      slope = computeSlope(rawRange, scaledRange)
      intercept = computeIntercept(slope, rawRange, scaledRange)
      scaledValue = slope * value + intercept
      return clipScaledValue(scaledValue, scaledRange)
  end

  def limit(value, range):
      return scale(value, range, range)
  end


  rq_init_comm_if_connected(9, "1")
  rq_init_comm_if_connected(2, "2")
  rq_init_comm_if_connected(3, "3")
  rq_init_comm_if_connected(4, "4")
  rq_print_connected_grippers()
  rq_gripper_communication_thread = run rq_gripper_communication()
  set_closed_norm(97.6470588235294, 1)
  set_open_norm(1.1764705882352942, 1)
  set_closed_mm(0.0, 1)
  set_open_mm(53.0, 1)
  set_closed_norm(100.0, 2)
  set_open_norm(0.0, 2)
  set_closed_mm(0.0, 2)
  set_open_mm(50.0, 2)
  set_closed_norm(100.0, 3)
  set_open_norm(0.0, 3)
  set_closed_mm(0.0, 3)
  set_open_mm(50.0, 3)
  set_closed_norm(100.0, 4)
  set_open_norm(0.0, 4)
  set_closed_mm(0.0, 4)
  set_open_mm(50.0, 4)
  rq_current_limit_enabled = False
  while(not rq_gripper_communication_thread_started):
      sync()
  end
  # end: URCap Installation Node
  # begin: URCap Installation Node
  #   Source: OPC UA, 2.0.2, Rocketfarm AS
  #   Type: OPC UA
  global opcua_daemon = rpc_factory("xmlrpc", "http://127.0.0.1:40409/RPC2")
  def opcua_client_connect(address):
  return opcua_daemon.client_connect(address)
  end
  def opcua_client_get_id(client_name):
  return opcua_daemon.client_get_id(client_name)
  end
  def opcua_client_try_connect(client_id):
  opcua_result = False
  if (opcua_daemon.client_connect(client_id)):
  sleep(0.01)
  opcua_result = opcua_daemon.client_is_connected(client_id)
  opcua_retry = 10
  while ( (not opcua_result) and (opcua_retry > 0) ):
  sleep(0.1)
  opcua_result = opcua_daemon.client_is_connected(client_id)
  opcua_retry = opcua_retry - 1
  end
  end
  return opcua_result
  end
  def opcua_client_disconnect(client_id):
  return opcua_daemon.client_disconnect(client_id)
  end
  def opcua_client_is_connected(client_id):
  return opcua_daemon.client_is_connected(client_id)
  end
  def opcua_client_read_byid(client_id, namespace_id, variable_id):
  return opcua_daemon.client_read_variable_by_id(client_id, namespace_id, variable_id)
  end
  def opcua_client_read_byname(client_id, namespace_id, variable_name):
  return opcua_daemon.client_read_variable_by_name(client_id, namespace_id, variable_name)
  end
  def opcua_client_write_byid(client_id, namespace_id, variable_id, variable_value):
  return opcua_daemon.client_write_variable_by_id(client_id, namespace_id, variable_id, variable_value)
  end
  def opcua_client_write_byname(client_id, namespace_id, variable_name, variable_value):
  return opcua_daemon.client_write_variable_by_name(client_id, namespace_id, variable_name, variable_value)
  end
  def opcua_client_last_error(client_id):
  return opcua_daemon.client_get_last_error(client_id)
  end
  def opcua_server_read_byname(variable_name):
  return opcua_daemon.server_read_variable_by_name(variable_name)
  end
  def opcua_server_write_byname(variable_name, variable_value):
  return opcua_daemon.server_write_variable_by_name(variable_name, variable_value)
  end
  def opcua_server_last_error():
  return opcua_daemon.server_get_last_error()
  end
  def opcua_error_to_string(errorCode):
  return opcua_daemon.error_code_to_string(errorCode)
  end
  # end: URCap Installation Node
  global AMR_Position=struct(position_identifier=0, x1=0, x2=0, y1=0, y2=0, theta1=0, theta2=0)
  global CAM_Pose=p[0,0,0,0,0,0]
  global CAM_Relation=""
  global CMD_Abort=  False
  global CMD_Clear=  False
  global CMD_Reset=  False
  global CMD_Start=  False
  global CMD_Suspend=  False
  global CMD_Unhold=  False
  global CMD_Unsuspend=  False
  global CNT_Rack_Output=0
  global FNC_Freedrive=  False
  global PRC_TubCounter=0
  global STP=0
  global easyPickCount=0
  global easyPickCount_4=0
  global easyPickCount_6=0
  global easyPickNoObj=0
  global easyPickNoObj_4=0
  global easyPickNoObj_6=0
  global easyPickParts=0
  global easyPickParts_4=0
  global easyPickParts_6=0
  global Container_mid_1_p=p[-.379239199143, -.127191311915, .299999999998, .000000000046, -.000000000021, -1.247199999994]
  global Container_mid_1_q=[-2.477408934449926, -1.2969853503591224, -1.875639182904262, -1.539621866126728, 1.5731943360401213, -2.8009955944022717]
  global Container_capt_p=p[-.525590029047, .407247642794, .411588185841, -.000000000107, .000000000065, -2.896148821900]
  global Container_capt_q=[-3.5968351615224767, -2.0050156108707204, -0.8176271154495112, -1.8895759482008394, 1.5730967555598792, -2.2743681102957645]
  global Waypoint_51_p=p[-.335468094724, -.217855817953, .299999999998, .000000000047, -.000000000014, -.994837065669]
  global Waypoint_51_q=[-2.2250460001249586, -1.2969853503591224, -1.875639182904262, -1.539621866126728, 1.573194336040121, -2.800995594402271]
  global Waypoint_65_p=p[-.380578560601, .136229906820, .300065486591, .002668209125, -.001950299791, -1.918285884015]
  global Waypoint_65_q=[-3.1484482924090784, -1.309784547691681, -1.8656262159347534, -1.5396564540318032, 1.5732260942459106, -2.8009706179248255]
  global Waypoint_86_p=p[-.610891912545, .328076512140, .154928874949, -.144389774448, 2.158207980619, -2.101916875088]
  global Waypoint_86_q=[-3.0298424402820032, -2.1616608105101527, -1.770405888557434, -1.8800016842284144, -0.04927570024599248, -0.4936583677874964]
  global Waypoint_16_p=p[-.530358413935, .418971000515, -.109643658887, -.463059997969, 2.087871459122, -2.058033430549]
  global Waypoint_16_q=[-3.2300904432879847, -2.6409207783141078, -1.877760410308838, -1.6937691173949183, -0.43063193956484014, 0.029483795166015625]
  global Waypoint_87_p=p[-.459488806274, .188986755628, .171097942578, -.348072585494, -2.059579317749, 2.019661285019]
  global Waypoint_87_q=[-2.790591303502218, -2.152559896508688, -1.6884642839431763, -2.469414850274557, 0.6884214878082275, 0.021232735365629196]
  global Waypoint_89_p=p[-.261886355761, -.111669623901, .131097242659, -1.173634433322, -1.227274747052, 1.193766216763]
  global Waypoint_89_q=[-2.672995464666928, -2.175407175402028, -1.7617490112425536, -2.338843663300132, 2.030865036219133, 0.036428578240585985]
  global Waypoint_90_p=p[-.269165142951, -.108082457315, .026677271969, -1.173634433324, -1.227274747052, 1.193766216762]
  global Waypoint_90_q=[-2.6853380119023815, -2.380020912479904, -1.7522585114443245, -2.1436252765786143, 2.018787725064888, 0.03659425986402358]
  global Waypoint_88_p=p[-.617446503519, .392270291627, .170489198955, -.224010410006, -2.066036920971, 2.088909130040]
  global Waypoint_88_q=[-3.1488035953258766, -2.4221038789008897, -1.1666724558911366, -2.618578428321003, 0.2380794033913185, -0.04528854192806264]
  global Waypoint_94_p=p[-.452978066378, .173533334300, .109390198136, -.002578830757, -2.196586508502, 2.177068753404]
  global Waypoint_94_q=[-2.6674557574892073, -2.1212895090252317, -1.967198705482553, -2.208419381150989, 0.5117897724834828, 0.04481344519449531]
  global Waypoint_93_p=p[-.596468537907, .142788156334, .105779109453, -.673355127215, 1.831389627653, -1.853156743314]
  global Waypoint_93_q=[-2.6921545586066635, -2.073966887503291, -2.065600898968258, -2.154852607781155, -0.22224352987151796, 0.042304121657345886]
  global Waypoint_95_p=p[-.605386387448, -.069660570533, .218481828695, .000812734400, .006677866481, -1.958478278110]
  global Waypoint_95_q=[-2.8029143834677903, -1.8400819882842256, -1.544169955118452, -1.327224466208456, 1.5676652012497132, -2.4155226342256775]
  global Waypoint_13_p=p[-.479450777041, .284140798427, .125270103493, -.276792173670, 2.098433187455, -2.121256516887]
  global Waypoint_13_q=[-2.8915050665484827, -1.9549266300597132, -2.2318272590637207, -1.6654960117735804, 0.020810842514038086, -0.4019392172442835]
  global Waypoint_70_p=p[-.472820924464, .292439826304, .207418370234, -.259787347864, -2.053484648504, 2.070709755662]
  global Waypoint_70_q=[-2.969927421603815, -2.07168115810532, -1.6835546062719366, -2.4953958198513964, 0.4489790927922641, -0.005578998612037367]
  global Waypoint_2_p=p[-.312961047461, -.152991312519, .223609826854, -.745314530454, -1.713873240489, 1.673341715282]
  global Waypoint_2_q=[-2.3560472170459192, -2.183784624139303, -1.4583134651184082, -2.6435262165465296, 1.6522362232208252, 0.043451953679323196]
  global Waypoint_3_p=p[-.113749865836, -.390110151572, .317307487562, -.519383711706, -.839884211339, 1.756868173041]
  global Waypoint_3_q=[-1.8909733931170862, -1.720626016656393, -1.5115610361099243, -2.1240560017027796, 2.1809096336364746, 0.7227501273155212]
  global Waypoint_15_p=p[.029144035010, -.436802470887, .327885032028, -.521560953301, -.623641814548, 1.862659450154]
  global Waypoint_15_q=[-1.564817253743307, -1.556895188321807, -1.6826975345611572, -1.6944714985289515, 2.2362685203552246, 1.117417335510254]
  global Waypoint_14_p=p[.068712235638, -.569419545175, .285215357659, -.679242949116, -.712065334485, 1.394044574094]
  global Waypoint_14_q=[-1.5731792953485346, -1.8029235103747094, -1.6781008808776736, -1.2218450646111982, 2.4719572998240125, 1.6394218026856375]
  global Waypoint_4_p=p[-.047220457210, -.557624911767, .136370962514, -.679242949107, -.712065334475, 1.394044574096]
  global Waypoint_4_q=[-1.7740079055958748, -2.0023561428872334, -1.7577251142892676, -1.18903287716154, 2.4487287370345143, 1.322902469273079]
  global Waypoint_25_p=p[.065436479647, -.569388431626, .287820755049, -.679242949185, -.712065334557, 1.394044574070]
  global Waypoint_25_q=[-1.5789263550890595, -1.8020194754825436, -1.6702557537748035, -1.237882536889547, 2.471995808083492, 1.6301087487321393]
  global Waypoint_39_p=p[.137772150180, -.577759956854, .299999999946, .000000000217, -.000000000207, -1.594351842625]
  global Waypoint_39_q=[-1.108978697428574, -1.776486680444405, -1.413737665315093, -1.5218908901738937, 1.5733062372356947, -1.0863866394180182]
  global Waypoint_41_p=p[.074222967010, -.565641640647, .234620140366, -.516884386806, .529223682286, -1.529619060506]
  global Waypoint_41_q=[-0.9596722604286052, -1.8767069964135548, -1.4892746174057256, -1.7813862040292285, 1.0520698599867686, -0.8199687448260349]
  global Waypoint_40_p=p[.039987741677, -.564832865048, .191055405868, -.767560686167, .343136533060, -2.241315728308]
  global Waypoint_40_q=[-1.0070649180116558, -1.8745927522477324, -1.6139175023195245, -1.6337474788493545, 1.032708081143138, -0.11587278312988403]
  global Waypoint_42_p=p[.041363380882, -.564865360786, .192805844739, .278500165520, .624117100927, .762272396553]
  global Waypoint_42_q=[-1.0050718976263102, -1.8744386685524779, -1.609151451954446, -1.6399653140247947, 1.0334006002355505, -3.254032861659603]
  global Waypoint_43_p=p[.041363380886, -.564865360780, .192805844755, .854271020883, .226833028600, 2.453002871494]
  global Waypoint_43_q=[-1.0050567614299233, -1.874341297657562, -1.6092945416026048, -1.6397580431809713, 1.0333661149462194, -5.0371728933995605]
  global Waypoint_44_p=p[.040882892233, -.564854254876, .192193763716, .110913882012, .659173708659, .275719738520]
  global Waypoint_44_q=[-1.0057704811530535, -1.8745207681598055, -1.6107765025572558, -1.637858394640876, 1.033164860873599, -2.7487836132940755]
  global Waypoint_45_p=p[.042647731639, -.564895808997, .194439423694, -.451694728506, .563172064821, -1.343350300184]
  global Waypoint_45_q=[-1.0032860829914387, -1.8741561795270565, -1.6048483308761785, -1.6453689714776623, 1.0342050634514657, -1.06078829880322]
  global Waypoint_46_p=p[.099944144487, -.566244126804, .267342790130, -.451694834765, .563172023386, -1.343350532536]
  global Waypoint_46_q=[-0.9257438092434924, -1.889970530402497, -1.3828165217629076, -1.8916791100652528, 1.0664350961373816, -0.9805910833329659]
  global Waypoint_47_p=p[.099944144444, -.566244126727, .267342790273, -.101742139519, .058679218003, -1.457888523314]
  global Waypoint_47_q=[-1.1112623176383014, -1.729989471869196, -1.5530029871033957, -1.4442770617454777, 1.4670579052775654, -1.2224020460061675]
  global Waypoint_48_p=p[-.136182767566, -.647487115908, .294247768372, -.101742139549, .058679218020, -1.457888523312]
  global Waypoint_48_q=[-1.532196177857717, -1.9115932455375173, -1.2651848069729779, -1.5055651746702665, 1.4703193777418382, -1.646379689188814]
  global Waypoint_49_p=p[-.159024328559, -.641021381179, .047691706070, -.000000000033, -.000000000027, -1.457897102937]
  global Waypoint_49_q=[-1.6098490079965062, -2.1164987141784586, -1.6156631902166785, -0.9800092198841526, 1.573231151532669, -1.722204302767242]
  global Waypoint_50_p=p[-.159024328558, -.641021381151, .291114489351, -.000000000033, -.000000000027, -1.457897102937]
  global Waypoint_50_q=[-1.609190265995684, -1.9426985888940234, -1.2189094859258596, -1.55056435122874, 1.5734384912955113, -1.7235116759964022]
  global Waypoint_53_p=p[-.050111345339, -.357608435610, .335880801283, .034180375734, .020280946727, -.284888945062]
  global Waypoint_53_q=[-1.3262308189700454, -1.2221767968893875, -1.8246061249803773, -1.7046285947349489, 1.567288986353525, -2.612420684434543]
  global Spatula_above_p=p[.240417564690, -.250827350286, .422801778001, .000126133258, .000019566993, -.045497134322]
  global Spatula_above_q=[-0.4110710190165463, -1.2060566172281924, -1.6172668714852705, -1.8889350758294619, 1.573016581809478, -1.9375501213280995]
  global Spatula_pick_p=p[.245838473482, -.255593930771, .230843335453, .000126133133, .000019564704, -.045497134323]
  global Spatula_pick_q=[-0.4194386807260848, -1.1902770326089298, -2.122244212434893, -1.399738227295769, 1.573431592600495, -1.943921578313585]
  global container_start_p=p[.200650292946, -.570238751958, .366326773614, 1.360500828661, .021700128770, 2.681649891414]
  global container_start_q=[-0.7669977765142582, -2.188996679669204, -0.7412727239230232, -2.581362891432544, 1.0193601740278728, 1.1884911920528847]
  global container_wp_1_p=p[.170613637794, -.572150573676, .294509026043, 1.259497117139, -.008270589399, 2.787717865625]
  global container_wp_1_q=[-0.8129253370121727, -2.0726598902108755, -1.0846040680899218, -2.2403146195823957, 1.0281191187839607, 1.0435744211830564]
  global Waypoint_55_p=p[.077280900603, -.567308602990, .212067617714, 1.259497117148, -.008270589399, 2.787717865619]
  global Waypoint_55_q=[-0.9181858327853867, -1.9744793804952083, -1.4540279077890048, -1.9155621911627945, 0.9643238328181578, 0.9457250675800015]
  global Waypoint_56_p=p[.135568164031, -.570867938153, .245215470413, 1.476861317558, -.018269607491, 2.679642659499]
  global Waypoint_56_q=[-0.8259784040282607, -2.108036981522602, -1.2111990877342924, -2.2405969375728745, 0.9451797152137279, 1.125710531287379]
  global Waypoint_74_p=p[.164827890887, -.574638012411, .193751361296, 2.053636896063, -.046507887560, 2.274278266449]
  global Waypoint_74_q=[-0.7657213433975762, -2.450387120010788, -0.9886183070290357, -2.7078095590939375, 0.8831550681477878, 1.5106229631053527]
  global ftr_scoop2_p=p[.194287054614, -.495779761333, .282072128495, -.179029871953, 1.612108092436, -.016025695011]
  global ftr_scoop2_q=[-0.5957383150173561, -2.264100500923713, -1.1936887184643812, -2.8893702964346097, 0.8750688478879766, -1.4109843517598684]
  global aftr_scoo3_p=p[-.289759911340, -.315385007342, .303743796282, .159961590809, 1.627415489603, -.344855744095]
  global aftr_scoo3_q=[-1.3374747909924949, -1.6809733407851706, -1.9857606509106667, -2.713564895186775, 0.5589807453366573, -1.3631067603374376]
  global Waypoint_60_p=p[-.013316432876, -.544772031582, .383371643081, 2.208233379808, .037543335712, 2.097559881761]
  global Waypoint_60_q=[-0.9328326161883087, -2.0999933666355775, -1.1958015693111372, -3.060905141293654, 0.690378518537611, 1.7121940951337198]
  global Waypoint_61_p=p[-.412188693372, -.356446875193, .383371643081, 1.751740964455, -.739956256289, 1.600691174920]
  global Waypoint_61_q=[-1.766185342973321, -2.0999933666355775, -1.1958015693111372, -3.060905141293654, 0.690378518537611, 1.7121940951337198]
  global Waypoint_75_p=p[-.343126484123, -.342779621892, .335357223804, .359429517288, 1.600352990741, -.365083732359]
  global Waypoint_75_q=[-1.517806275013295, -1.8136828056045395, -1.737638081810795, -2.8432599585466436, 0.5149430839716123, -1.4579122147201877]
  global aftr_scoop1_p=p[.138503854266, -.514479969882, .214153672011, -.134825326227, 1.559916297527, -.059196589314]
  global aftr_scoop1_q=[-0.6880464314785328, -2.2689986529709643, -1.3310176475983653, -2.673087158390708, 0.8340516295138949, -1.4557846480003231]
  global After_disp_3_p=p[.125934854156, -.585611107804, .299545938076, .959554236104, -.134386766509, 2.880651774211]
  global After_disp_3_q=[-0.9434480594885066, -2.016473586333989, -1.1036579072158617, -2.096459283015281, 1.1479556364931514, 0.8433331387406042]
  global Waypoint_62_p=p[-.542658707241, -.114281911009, .251261544113, 1.813043609523, -.679411528034, 1.655271622964]
  global Waypoint_62_q=[-2.158300033470912, -1.9418836862428677, -1.8142999147147894, -2.778920736683023, 0.21900622104017292, 1.8983390235012934]
  global Waypoint_63_p=p[.101294795191, -.465376052375, .381756220355, .972633305146, -.158447626639, 2.887199602585]
  global Waypoint_63_q=[-0.8528172446194038, -1.7393709485118478, -1.2544079521837954, -2.2703112963960628, 1.1965892397133469, 0.91867216443391]
  global Start_p=p[-.033064633790, -.365398531763, .389873206922, .000000000001, .000000000001, 2.725785203584]
  global Start_q=[-1.287596562866887, -1.232866726886848, -1.6880113260231102, -1.7912103151657988, 1.5729028131945846, 0.6981423183093938]
  global Waypoint_76_p=p[-.479450777041, .284140798427, .125270103493, -.276792173670, 2.098433187454, -2.121256516887]
  global Waypoint_76_q=[-2.891505066548503, -1.9549266300590151, -2.231827259067863, -1.6654960117542226, 0.020810842514162875, -0.4019392172601952]
  global PowderA_wayp1_p=p[-.472820924474, .292439826233, .207418370237, -.137787250486, 2.177332259632, -2.152029714756]
  global PowderA_wayp1_q=[-2.911134078210732, -1.90240864358569, -1.968768330510411, -2.500365101593811, 0.11427687110891149, 0.0958980389250167]
  global Waypoint_80_p=p[-.303921889165, -.326082520111, .297721580072, -.584846481381, 1.914382606328, -1.960922301253]
  global Waypoint_80_q=[-1.6364180099980672, -2.041258366871811, -1.472153549517767, -2.7572808013122696, 0.9684003593854582, 0.047163023020230455]
  global Decapp_above_p=p[-.013480295948, -.359153355979, .266194408367, -.879653555922, 1.646336924805, -1.709111068605]
  global Decapp_above_q=[-0.9632157249872035, -2.0163405763031657, -1.5968194594157152, -2.6579215719847085, 1.251243398585566, 0.047906446502667066]
  global Decapp_place_p=p[-.013480295848, -.359153356116, .158558645017, -.879653554904, 1.646336919751, -1.709111066446]
  global Decapp_place_q=[-0.9633419174801583, -2.157735564881908, -1.695182597572722, -2.418253553201909, 1.2517436353048952, 0.04819090596102882]
  global Waypoint_78_p=p[-.051450028091, -.519555688329, .365718563414, -1.287302938145, 1.077637394477, -1.218524965834]
  global Waypoint_78_q=[-0.9214276262416012, -1.8899696965062578, -1.4939326452510562, -2.840015661555725, 0.5585157189668353, 0.033997638875617575]
  global Waypoint_81_p=p[-.030847790230, -.346237542439, .241203613248, .000000000000, .000000000000, .000000000000]
  global Waypoint_81_q=[-1.265848516232941, -1.1652881302267932, -2.11003646605462, -1.4369228603041853, 1.573284436504383, -2.835929896730388]
  global Waypoint_79_p=p[-.030847972829, -.346235312674, .229874122470, .000000000000, .000000000000, .000000000000]
  global Waypoint_79_q=[-1.2659333103898618, -1.1699230683425625, -2.1365870669440055, -1.4057372655396474, 1.5732787836040316, -2.8358953794066757]
  global Waypoint_82_p=p[-.031079593487, -.346547394534, .293012696855, -.000011575267, -.000017731224, -.000713984074]
  global Waypoint_82_q=[-1.2664169521879751, -1.1572597700415788, -1.982185304253158, -1.5727862504184884, 1.5732673022058234, -2.83632822711502]
  global Cap_above_p=p[-.163602500478, -.618357694237, .258271116068, .000026793591, -.000032305852, -.969382601663]
  global Cap_above_q=[-1.6181634639269902, -1.896432778341337, -1.3662765317923142, -1.449515114018281, 1.5734416863575176, -2.220489512402157]
  global Cap_Place_p=p[-.153420247224, -.637174247221, .035295616791, .000000000002, -.000000000002, -1.457849918374]
  global Cap_Place_q=[-1.6014084627078784, -2.123124488207292, -1.6429187572395012, -0.946127085055064, 1.573175527437006, -1.7136981844648291]
  global OP_PowderA2_p=p[.009371277507, -.409434369247, .294169017766, -.823281033205, 1.709410851243, -1.698303593897]
  global OP_PowderA2_q=[-0.9994544761745754, -2.1395254572673217, -1.3437567783153916, -2.8143375616690456, 1.2617899549595724, 0.019614613715634555]
  global OP_PowderA_abov_p=p[-.012145216791, -.363335041455, .315325728178, -.777135478411, 1.752984823781, -1.740925591659]
  global OP_PowderA_abov_q=[-1.01634425044037, -2.024785947780374, -1.4658894155189923, -2.8070189735738786, 1.3091674480404514, 0.020022086766872782]
  global OP_PowderA_pick_p=p[-.012145216707, -.363335041590, .179898787547, -.777135478413, 1.752984823781, -1.740925591659]
  global OP_PowderA_pick_q=[-1.0165129229305911, -2.176980100858497, -1.6127054339661555, -2.5080740815244567, 1.3098787614888208, 0.020270375244195882]
  global Tilt_above_p=p[-.111064400266, -.518714782683, .336190805493, -1.186264705469, 1.271052138367, -1.268665700837]
  global Tilt_above_q=[-1.0593782044036235, -1.983218206819794, -1.4684292238819445, -2.8468741750118465, 0.5899608864573523, 0.021166292918283425]
  global Tilt_place_p=p[-.116477368770, -.516998826303, .220965575609, -1.186264705477, 1.271052138372, -1.268665700834]
  global Tilt_place_q=[-1.0667718212381487, -2.0926346913000655, -1.6256300657432945, -2.5807129872023205, 0.5834128338282412, 0.021733786155414034]
  global Waypoint_52_p=p[-.141928460719, -.515782557948, .252798475575, .000000001021, .000000015714, -1.648489523537]
  global Waypoint_52_q=[-1.5865298660227536, -1.6477298798514424, -1.683499112918053, -1.3809236418182405, 1.5732592408189925, -1.5089407655972176]
  global ViaPoint_1_p=p[-.075380379718, -.518346610957, .240267869004, -.308187611455, .314849234097, -1.629298408213]
  global ViaPoint_1_q=[-1.2665498468402658, -1.632968153584656, -1.7466488267795093, -1.4757122352125567, 1.206407674916738, -1.1583391815257933]
  global Waypoint_57_p=p[-.016929050533, -.520720414258, .208138086750, -.566600031366, .578847302089, -1.576463827532]
  global Waypoint_57_q=[-1.0408435604305932, -1.753222942634757, -1.738239877480245, -1.6732057965873945, 0.9875721214075002, -0.8174462985078907]
  global Waypoint_69_p=p[.038244169892, -.523681622326, .270660553693, -.566600038239, .578847306557, -1.576463843233]
  global Waypoint_69_q=[-0.9584046232102423, -1.7662930703212236, -1.5465420531532832, -1.8980111501412296, 1.0250918773452096, -0.7315432464998608]
  global PowA_ScoopA_p=p[.159611615818, -.500668442765, .327719041452, -.697225816707, .808151787064, -1.272841262549]
  global PowA_ScoopA_q=[-0.7052336156646533, -1.9354458065172322, -1.2435429111590262, -2.383130756765686, 0.9889263119369867, -0.6132400042961272]
  global scoop_p=p[.074657261350, -.519131732172, .256549412299, -.011051468192, .988408833954, .005144340905]
  global scoop_q=[-0.8274053586011583, -1.874926877200366, -1.5200461069833828, -2.106983319332074, 0.9002119871547718, -2.116685021101622]
  global Waypoint_71_p=p[.177770645713, -.528015530173, .277526412330, .001909155730, 1.639086158711, -.035491055298]
  global Waypoint_71_q=[-0.6883155724662711, -2.3735431185097156, -1.0244077123914472, -2.9690624372933723, 0.9072837830600953, -1.4995275296364206]
  global Waypoint_83_p=p[.150765656890, -.528941996739, .207349351161, .001909146913, 1.639086162262, -.035491054401]
  global Waypoint_83_q=[-0.715557591216621, -2.395263074398475, -1.1745539289501714, -2.7990107897487184, 0.8808120190924962, -1.4964991406090151]
  global Waypoint_73_p=p[.145083518034, -.526977858919, .266012644295, -.001096606732, 1.243803685484, -.039558884435]
  global Waypoint_73_q=[-0.7315307126590884, -2.1222688412291646, -1.2371995036129686, -2.500626334721838, 0.9062275384215436, -1.820210419506548]
  global aftr_disp4_p=p[.076649091963, -.516683659078, .327659997949, -.089442013925, .747027934620, -.179429504000]
  global aftr_disp4_q=[-0.8729541889129182, -1.7538731498931135, -1.421722565562387, -2.0624433405073983, 1.0093695837082866, -2.1021195561352615]
  global Waypoint_84_p=p[.123174711194, -.515520147762, .377487231436, -.089442013731, .747027928699, -.179429504004]
  global Waypoint_84_q=[-0.8099995125927881, -1.8159482911699527, -1.2110272502558486, -2.243587231698566, 1.0414314296112155, -2.0397317655088933]
  global Waypoint_54_p=p[.127020102667, -.520474555499, .444734866371, -.000000000049, -.000000000029, -.181836163636]
  global Waypoint_54_q=[-1.077914415145683, -1.67713376904155, -1.1559751108552438, -1.8791222047311322, 1.5728513980826264, -2.469046273458339]
  global Waypoint_58_p=p[.222355978426, -.256721511160, .377517216113, .000126133135, .000019564704, -.045497133314]
  global Waypoint_58_q=[-0.4523685080439055, -1.1582470295698233, -1.764486450044644, -1.7895331365539002, 1.573203470967134, -1.9783680221047675]
  global Waypoint_59_p=p[.246090929453, -.257346948962, .334937874481, .002062251865, .085969144325, -.045466267072]
  global Waypoint_59_q=[-0.3993250128175445, -1.229937207675869, -1.8134849075269486, -1.7494730648138157, 1.5434956294817688, -1.9239935269750585]
  global Waypoint_72_p=p[.241373394141, -.257127682308, .280144245911, .002062251870, .085969144324, -.045466267071]
  global Waypoint_72_q=[-0.40453618428666793, -1.2163524390607545, -1.961899201118312, -1.614505550067273, 1.54321918600584, -1.9286199875396806]
  global Waypoint_68_p=p[-.054140750939, -.519225939047, .230771617164, -.396603942010, .405176681937, -1.615073614845]
  global Waypoint_68_q=[-1.1801200722220573, -1.66078878572511, -1.7519948628362751, -1.5321103532497595, 1.1202658922042295, -1.0435495794713274]
  global Waypoint_67_p=p[-.085538600094, -.517926057057, .244809615848, -.265837410279, .271583584295, -1.634720190296]
  global Waypoint_67_q=[-1.3101477871233094, -1.6246275760972235, -1.7396885526482375, -1.4554188629779246, 1.2515887427265664, -1.211612237682651]
  global Waypoint_66_p=p[-.112404525053, -.516834057197, .249908478866, -.145067433961, .148203121183, -1.645288419275]
  global Waypoint_66_q=[-1.4361046238427022, -1.62151199833529, -1.7216739172895004, -1.4033237867418515, 1.391749278833954, -1.3534436213375054]
  global Waypoint_77_p=p[-.029562189306, -.345402935881, .227061086376, -.000128098079, -.000007607820, -.000007077939]
  global Waypoint_77_q=[-1.2613241377464561, -1.168338291946169, -2.144792803677632, -1.3989918632055023, 1.5732473641903764, -2.831248128197144]
  def Sub_Vision_V18():
    $ 672 "Sub_Vision_V18" "noBreak"
    $ 673 "PreSettings"
    $ 674 "CAM_LM_Detected≔ False "
    global CAM_LM_Detected=  False
    $ 675 "CAM_Captures≔0"
    global CAM_Captures=0
    $ 676 "CAM_Pose≔p[0,0,0,0,0,0]"
    global CAM_Pose=p[0,0,0,0,0,0]
    $ 677 "CAM_LM_Refinmnt≔ False "
    global CAM_LM_Refinmnt=  False
    $ 678 "CAM_LM_Refined≔ False "
    global CAM_LM_Refined=  False
    $ 679 "CAM_LM_Deviatn≔p[0,0,0,0,0,0]"
    global CAM_LM_Deviatn=p[0,0,0,0,0,0]
    $ 680 "CAM_LM_ID≔0"
    global CAM_LM_ID=0
    $ 681 "CAM_Done≔ False "
    global CAM_Done=  False
    $ 682 "CAM_CNT_Obj≔0"
    global CAM_CNT_Obj=0
    $ 683 "CAM_Result = []"
    CAM_Result = []
    $ 684 "OBJ_Detected≔ False "
    global OBJ_Detected=  False
    $ 685 "FRM_Reference≔p[0,0,0,0,0,0]"
    global FRM_Reference=p[0,0,0,0,0,0]
    $ 686 "'=========='"
    # '=========='
    $ 687 "Switch Action"
    switch_1 = Action
    $ 688 "Case 13"
    if (13 == switch_1):
    elif (15 == switch_1):
      $ 806 "Case 15"
    elif (131 == switch_1):
      $ 852 "Case 131"
      $ 853 "Read (SensoPart)"
      $ 854 "Action_Info≔'search for landmark'"
      global Action_Info="search for landmark"
      $ 855 "CAM_LM≔CAM_LMs[4]"
      global CAM_LM=CAM_LMs[4]
      $ 856 "CAM_Relation≔CAM_LM.capture_relation"
      global CAM_Relation=CAM_LM.capture_relation
      $ 857 "go to capture pose"
      $ 860 "If ITM_ID≟1 and JIG≟7"
      if (ITM_ID == 1  and  JIG == 7):
        $ 861 "PSE_T≔uLM_Cap_SSRack"
        global PSE_T=uLM_Cap_SSRack
      else:
        $ 862 "ElseIf ITM_ID≟5 and JIG≟7"
        if (ITM_ID == 5  and  JIG == 7):
          $ 863 "PSE_T≔FRM_Cap_SSRack"
          global PSE_T=FRM_Cap_SSRack
        else:
          $ 864 "ElseIf ITM_ID≟13 and JIG≟7"
          if (ITM_ID == 13  and  JIG == 7):
            $ 865 "PSE_T≔FRM_pick_rack_const"
            global PSE_T=p[-0.5568395192387274,0.34423986364170267,0.44698620470146266,-1.0069110132199915E-6,3.378712467497258E-5,-8.002029546773325E-6]
          else:
            $ 866 "ElseIf ITM_ID≟1 and JIG≟15"
            if (ITM_ID == 1 and JIG == 15):
              $ 867 "MoveJ"
              $ 868 "Container_mid_1" "breakAfter"
              movej(get_inverse_kin(Container_mid_1_p, qnear=Container_mid_1_q), a=1.3962634015954636, v=1.0471975511965976, r=0.05)
              $ 869 "Container_capt" "breakAfter"
              movej(get_inverse_kin(Container_capt_p, qnear=Container_capt_q), a=1.3962634015954636, v=1.0471975511965976)
              $ 870 "PSE_T≔FRM_Container_S_const"
              global PSE_T=p[-0.510412665574981,0.40064363362973565,0.41159789496794374,-1.1370875604168537E-5,-3.643547521609506E-6,-2.896122366208473]
            else:
              $ 871 "ElseIf ITM_ID≟1 and JIG≟16"
              if (ITM_ID == 1  and  JIG == 16):
                $ 872 "MoveJ"
                $ 873 "Waypoint_51" "breakAfter"
                movej(get_inverse_kin(Waypoint_51_p, qnear=Waypoint_51_q), a=1.3962634015954636, v=1.0471975511965976, r=0.05)
                $ 876 "PSE_T≔FRM_Container_S_const"
                global PSE_T=p[-0.510412665574981,0.40064363362973565,0.41159789496794374,-1.1370875604168537E-5,-3.643547521609506E-6,-2.896122366208473]
              else:
                $ 877 "ElseIf ITM_ID≟1 and JIG≟17"
                if (ITM_ID == 1  and  JIG == 17):
                  $ 878 "MoveJ"
                  $ 879 "Waypoint_51" "breakAfter"
                  movej(get_inverse_kin(Waypoint_51_p, qnear=Waypoint_51_q), a=1.3962634015954636, v=1.0471975511965976, r=0.05)
                  $ 882 "PSE_T≔FRM_Container_S_const"
                  global PSE_T=p[-0.510412665574981,0.40064363362973565,0.41159789496794374,-1.1370875604168537E-5,-3.643547521609506E-6,-2.896122366208473]
                else:
                  $ 883 "ElseIf ITM_ID≟1 and JIG≟18"
                  if (ITM_ID == 1  and  JIG == 18):
                    $ 886 "MoveJ"
                    $ 887 "Waypoint_51" "breakAfter"
                    movej(get_inverse_kin(Waypoint_51_p, qnear=Waypoint_51_q), a=1.3962634015954636, v=1.0471975511965976, r=0.05)
                    $ 888 "Waypoint_65" "breakAfter"
                    movej(get_inverse_kin(Waypoint_65_p, qnear=Waypoint_65_q), a=1.3962634015954636, v=1.0471975511965976)
                    $ 889 "PSE_T≔FRM_Container_S_const"
                    global PSE_T=p[-0.510412665574981,0.40064363362973565,0.41159789496794374,-1.1370875604168537E-5,-3.643547521609506E-6,-2.896122366208473]
                  else:
                    $ 890 "ElseIf ITM_ID≟1 and JIG≟19"
                    if (ITM_ID == 1  and  JIG == 19):
                      $ 893 "MoveJ"
                      $ 894 "Waypoint_51" "breakAfter"
                      movej(get_inverse_kin(Waypoint_51_p, qnear=Waypoint_51_q), a=1.3962634015954636, v=1.0471975511965976, r=0.05)
                      $ 896 "PSE_T≔aq_rack1_const"
                      global PSE_T=p[-0.6171199234912242,0.18274496130308399,0.4990241423073791,7.867082192074154E-6,-3.513408957609815E-5,-2.5093516385827686]
                    end
                  end
                end
              end
            end
          end
        end
      end
      $ 897 "do_transition(PSE_T, keep_rxry=False)"
      do_transition(PSE_T, keep_rxry=False)
      $ 898 "Set"
      set_tcp(p[0.0,0.0,0.161,3.1415,0.0,0.0])
      $ 899 "MoveJ"
      $ 900 "PSE_T" "breakAfter"
      movej(PSE_T, a=1.3962634015954636, v=1.7453292519943295)
      $ 901 "CAM_Pose≔get_actual_tcp_pose()"
      global CAM_Pose= get_actual_tcp_pose ()
      $ 902 "Loop  not CAM_Done and  not ERROR.FLAG and  not CMD_Stop"
      while (  not  CAM_Done  and    not  ERROR.FLAG  and    not  CMD_Stop):
        $ 903 "adjust capture pose"
        $ 904 "If CAM_LM_Detected and CAM_LM_Refinmnt"
        if (CAM_LM_Detected  and  CAM_LM_Refinmnt):
          $ 905 "PSE_T≔p[0,0,0.300,0,0,0]"
          global PSE_T=p[0,0,0.300,0,0,0]
          $ 906 "CAM_Pose≔PSE_T"
          global CAM_Pose=PSE_T
          $ 907 "If  not is_reachable(FRM_Reference,[PSE_T])"
          if (  not  is_reachable(FRM_Reference,[PSE_T])):
            $ 908 "Error"
            $ 909 "set_error(ERROR_POSE_NOT_REACHABLE)"
            set_error(ERROR_POSE_NOT_REACHABLE)
          end
          $ 910 "If  not ERROR.FLAG"
          if (  not  ERROR.FLAG):
            $ 911 "MoveJ"
            $ 912 "PSE_T" "breakAfter"
            set_tcp(p[0.0,0.0,0.161,0.0,0.0,0.0])
            movej(pose_trans(FRM_Reference, PSE_T), a=0.8726646259971648, v=1.3962634015954636)
            $ 913 "CAM_LM_Refined≔ True "
            global CAM_LM_Refined=  True
          end
        else:
          $ 914 "ElseIf  not CAM_LM_Detected and CAM_Captures>0"
          if (  not  CAM_LM_Detected  and  CAM_Captures>0):
            $ 915 "MoveL"
            $ 916 "If FRM_Reference≟p[0,0,0,0,0,0]"
            if (FRM_Reference == p[0,0,0,0,0,0]):
              $ 917 "PSE_T≔get_random_pose(pose_ref=CAM_Pose, mode='cubic', range_max=[0.150,0.150,0.015])"
              global PSE_T=get_random_pose(pose_ref=CAM_Pose, mode="cubic", range_max=[0.150,0.150,0.015])
            else:
              $ 922 "Else" "noBreak"
              $ 923 "PSE_T≔get_random_pose(pose_ref=CAM_Pose, mode='rotation', range_max=[10,10,0])"
              global PSE_T=get_random_pose(pose_ref=CAM_Pose, mode="rotation", range_max=[10,10,0])
              $ 924 "CAM_LM_Refined≔ True "
              global CAM_LM_Refined=  True
            end
            $ 925 "If get_inverse_kin_has_solution(pose_trans(FRM_Reference, PSE_T))"
            if (get_inverse_kin_has_solution( pose_trans (FRM_Reference, PSE_T))):
              $ 926 "Comment"
              # Comment
              $ 927 "PSE_T" "breakAfter"
              set_tcp(p[0.0,0.0,0.161,3.1415,0.0,0.0])
              movel(pose_trans(FRM_Reference, PSE_T), a=0.03, v=0.05)
            else:
              $ 928 "Else" "noBreak"
              $ 929 "'If random pose is out of reach, set the initial cam pose'"
              # 'If random pose is out of reach, set the initial cam pose'
              $ 930 "PSE_T≔CAM_Pose"
              global PSE_T=CAM_Pose
            end
          end
        end
        $ 931 "Wait: 2.0"
        sleep(2.0)
        $ 932 "trigger"
        $ 933 "If ITM_ID≟1 and JIG≟7"
        if (ITM_ID == 1  and  JIG == 7):
          # begin: URCap Program Node
          #   Source: SensoPart VISOR Robotic, 2.0.0, SensoPart Industriesensorik GmbH
          #   Type: VISOR Trigger
          $ 934 "# 1 VISOR Trigger"
          visor_changeJob(1, "Landmark_INVITE_2", 6000)
          visor_trigger(1, 6000, "arm")
          # end: URCap Program Node
        else:
          $ 935 "ElseIf ITM_ID≟5 and JIG≟7"
          if (ITM_ID == 5  and  JIG == 7):
            # begin: URCap Program Node
            #   Source: SensoPart VISOR Robotic, 2.0.0, SensoPart Industriesensorik GmbH
            #   Type: VISOR Trigger
            $ 936 "# 1 VISOR Trigger"
            visor_changeJob(1, "Landmark_INVITE_2", 6000)
            visor_trigger(1, 6000, "arm")
            # end: URCap Program Node
          else:
            $ 937 "ElseIf ITM_ID≟13 and JIG≟7"
            if (ITM_ID == 13  and  JIG == 7):
              # begin: URCap Program Node
              #   Source: SensoPart VISOR Robotic, 2.0.0, SensoPart Industriesensorik GmbH
              #   Type: VISOR Trigger
              $ 938 "# 1 VISOR Trigger"
              visor_changeJob(1, "Landmark_INVITE_2", 6000)
              visor_trigger(1, 6000, "arm")
              # end: URCap Program Node
            else:
              $ 939 "ElseIf ITM_ID≟1 and JIG≟15"
              if (ITM_ID == 1 and JIG == 15):
                # begin: URCap Program Node
                #   Source: SensoPart VISOR Robotic, 2.0.0, SensoPart Industriesensorik GmbH
                #   Type: VISOR Trigger
                $ 940 "# 1 VISOR Trigger"
                visor_changeJob(1, "PowderA", 6000)
                visor_trigger(1, 6000, "arm")
                # end: URCap Program Node
              else:
                $ 941 "ElseIf ITM_ID≟1 and JIG≟16"
                if (ITM_ID == 1 and JIG == 16):
                  # begin: URCap Program Node
                  #   Source: SensoPart VISOR Robotic, 2.0.0, SensoPart Industriesensorik GmbH
                  #   Type: VISOR Trigger
                  $ 942 "# 1 VISOR Trigger"
                  visor_changeJob(1, "Weigh_target", 6000)
                  visor_trigger(1, 6000, "arm")
                  # end: URCap Program Node
                else:
                  $ 943 "ElseIf ITM_ID≟1 and JIG≟17"
                  if (ITM_ID == 1 and JIG == 17):
                    # begin: URCap Program Node
                    #   Source: SensoPart VISOR Robotic, 2.0.0, SensoPart Industriesensorik GmbH
                    #   Type: VISOR Trigger
                    $ 944 "# 1 VISOR Trigger"
                    visor_changeJob(1, "Weigh_dispense", 6000)
                    visor_trigger(1, 6000, "arm")
                    # end: URCap Program Node
                  else:
                    $ 945 "ElseIf ITM_ID≟1 and JIG≟18"
                    if (ITM_ID == 1 and JIG == 18):
                      # begin: URCap Program Node
                      #   Source: SensoPart VISOR Robotic, 2.0.0, SensoPart Industriesensorik GmbH
                      #   Type: VISOR Trigger
                      $ 946 "# 1 VISOR Trigger"
                      visor_changeJob(1, "pick_rack", 6000)
                      visor_trigger(1, 6000, "arm")
                      # end: URCap Program Node
                    else:
                      $ 948 "ElseIf ITM_ID≟1 and JIG≟19"
                      if (ITM_ID == 1 and JIG == 19):
                        # begin: URCap Program Node
                        #   Source: SensoPart VISOR Robotic, 2.0.0, SensoPart Industriesensorik GmbH
                        #   Type: VISOR Trigger
                        $ 949 "# 1 VISOR Trigger"
                        visor_changeJob(1, "place_rack", 6000)
                        visor_trigger(1, 6000, "arm")
                        # end: URCap Program Node
                      end
                    end
                  end
                end
              end
            end
          end
        end
        $ 954 "TM_3D≔visor_partsFound(1)"
        global TM_3D= visor_partsFound (1)
        $ 955 "If TM_3D>0"
        if (TM_3D>0):
          $ 956 "CAM_LM_Detected≔ True "
          global CAM_LM_Detected=  True
          $ 957 "CAM_Captures≔0"
          global CAM_Captures=0
        else:
          $ 958 "Else" "noBreak"
          $ 959 "CAM_LM_Detected≔ False "
          global CAM_LM_Detected=  False
          $ 960 "CAM_Captures≔CAM_Captures+1"
          global CAM_Captures=CAM_Captures+1
        end
        $ 965 "result"
        $ 966 "If CAM_LM_Detected"
        if (CAM_LM_Detected):
          $ 967 "If (CAM_LM_Refinmnt and CAM_LM_Refined) or  not CAM_LM_Refinmnt"
          if ((CAM_LM_Refinmnt  and  CAM_LM_Refined)  or    not  CAM_LM_Refinmnt):
            $ 1025 "If ITM_ID≟1 and JIG≟7"
            if (ITM_ID == 1  and  JIG == 7):
              $ 1026 "CAM_LM_SSRack≔visor_getPose3d(1, 0)"
              global CAM_LM_SSRack= visor_getPose3d (1, 0)
            else:
              $ 1027 "ElseIf ITM_ID≟5 and JIG≟7"
              if (ITM_ID == 5  and  JIG == 7):
                $ 1028 "CAM_LM_SSRack≔visor_getPose3d(1, 0)"
                global CAM_LM_SSRack= visor_getPose3d (1, 0)
              else:
                $ 1029 "ElseIf ITM_ID≟13 and JIG≟7"
                if (ITM_ID == 13  and  JIG == 7):
                  $ 1030 "CAM_LM_Bott≔visor_getPose3d(1, 0)"
                  global CAM_LM_Bott= visor_getPose3d (1, 0)
                else:
                  $ 1031 "ElseIf ITM_ID≟1 and JIG≟15"
                  if (ITM_ID == 1 and JIG == 15):
                    $ 1032 "CAM_LM_Cont_S≔visor_getPose3d(1, 0)"
                    global CAM_LM_Cont_S= visor_getPose3d (1, 0)
                    $ 1033 "cont_img_pose≔get_actual_tcp_pose()"
                    global cont_img_pose= get_actual_tcp_pose ()
                  else:
                    $ 1034 "ElseIf ITM_ID≟1 and JIG≟16"
                    if (ITM_ID == 1 and JIG == 16):
                      $ 1035 "CAM_cont≔visor_getPose3d(1, 0)"
                      global CAM_cont= visor_getPose3d (1, 0)
                      $ 1036 "cont_img_pose≔get_actual_tcp_pose()"
                      global cont_img_pose= get_actual_tcp_pose ()
                    else:
                      $ 1037 "ElseIf ITM_ID≟1 and JIG≟17"
                      if (ITM_ID == 1 and JIG == 17):
                        $ 1038 "pose_rack_aq1≔visor_getPose3d(1, 0)"
                        global pose_rack_aq1= visor_getPose3d (1, 0)
                        $ 1039 "cont_img_pose≔get_actual_tcp_pose()"
                        global cont_img_pose= get_actual_tcp_pose ()
                      else:
                        $ 1040 "ElseIf ITM_ID≟1 and JIG≟18"
                        if (ITM_ID == 1 and JIG == 18):
                          $ 1041 "pose_rack_aq1≔visor_getPose3d(1, 0)"
                          global pose_rack_aq1= visor_getPose3d (1, 0)
                          $ 1042 "FRM_Container_S≔get_actual_tcp_pose()"
                          global FRM_Container_S= get_actual_tcp_pose ()
                        else:
                          $ 1043 "ElseIf ITM_ID≟1 and JIG≟19"
                          if (ITM_ID == 1 and JIG == 19):
                            $ 1044 "pose_rack_aq1≔visor_getPose3d(1, 0)"
                            global pose_rack_aq1= visor_getPose3d (1, 0)
                            $ 1045 "aq_rack1≔get_actual_tcp_pose()"
                            global aq_rack1= get_actual_tcp_pose ()
                          end
                        end
                      end
                    end
                  end
                end
              end
            end
            $ 1046 "CAM_Done≔ True "
            global CAM_Done=  True
          end
        else:
          $ 1047 "ElseIf  not CAM_LM_Detected and CAM_Captures<CAM_PRM_Retries"
          if (  not  CAM_LM_Detected  and  CAM_Captures<CAM_PRM_Retries):
            $ 1048 "CAM_LM_Refined≔ False "
            global CAM_LM_Refined=  False
          else:
            $ 1049 "ElseIf CAM_Captures≥CAM_PRM_Retries"
            if (CAM_Captures >= CAM_PRM_Retries):
              $ 1050 "CAM_Done≔ True "
              global CAM_Done=  True
              $ 1051 "Error"
              $ 1052 "set_error(ERROR_NO_LANDMARK)"
              set_error(ERROR_NO_LANDMARK)
            end
          end
        end
      end
    elif (151 == switch_1):
      $ 1053 "Case 151"
      $ 1054 "Detect (SensoPart)"
      $ 1055 "go to capture pose"
      $ 1056 "FRM_Reference≔FRM_Cap_SSRack"
      global FRM_Reference=FRM_Cap_SSRack
      $ 1057 "PSE_T≔p[0,0,-0.00,0,0,0]"
      global PSE_T=p[0,0,-0.00,0,0,0]
      $ 1058 "do_transition(pose_trans(FRM_Reference, PSE_T), keep_rxry=False)"
      do_transition( pose_trans (FRM_Reference, PSE_T), keep_rxry=False)
      $ 1059 "JNT_Q≔get_actual_joint_positions()"
      global JNT_Q= get_actual_joint_positions ()
      $ 1060 "JNT_Q≔[JNT_Q[0], JNT_Q[1], JNT_Q[2], JNT_Q[3], JNT_Q[4], 0]"
      global JNT_Q=[JNT_Q[0], JNT_Q[1], JNT_Q[2], JNT_Q[3], JNT_Q[4], 0]
      $ 1061 "Set"
      set_tcp(p[0.0,0.0,0.161,3.1415,0.0,0.0])
      $ 1062 "movej(get_inverse_kin(pose_trans(FRM_Reference, PSE_T), qnear=JNT_Q))"
      movej(get_inverse_kin( pose_trans (FRM_Reference, PSE_T), qnear=JNT_Q))
      $ 1063 "CAM_Pose≔pose_trans(pose_inv(FRM_Reference), get_actual_tcp_pose())"
      global CAM_Pose= pose_trans ( pose_inv (FRM_Reference),  get_actual_tcp_pose ())
      $ 1064 "Loop  not CAM_Done and  not ERROR.FLAG and  not CMD_Stop"
      while (  not  CAM_Done  and    not  ERROR.FLAG  and    not  CMD_Stop):
        $ 1065 "If  not OBJ_Detected and CAM_Captures>0"
        if (  not  OBJ_Detected  and  CAM_Captures>0):
          $ 1066 "MoveL"
          $ 1067 "If FRM_Reference≟p[0,0,0,0,0,0]"
          if (FRM_Reference == p[0,0,0,0,0,0]):
            $ 1069 "PSE_T≔get_random_pose(pose_ref=CAM_Pose, mode='rotation', range_max=[15,15,0])"
            global PSE_T=get_random_pose(pose_ref=CAM_Pose, mode="rotation", range_max=[15,15,0])
          else:
            $ 1070 "Else" "noBreak"
            $ 1071 "PSE_T≔get_random_pose(pose_ref=CAM_Pose, mode='rotation', range_max=[10,10,0])"
            global PSE_T=get_random_pose(pose_ref=CAM_Pose, mode="rotation", range_max=[10,10,0])
          end
          $ 1072 "If get_inverse_kin_has_solution(pose_trans(FRM_Reference, PSE_T))"
          if (get_inverse_kin_has_solution( pose_trans (FRM_Reference, PSE_T))):
            $ 1073 "PSE_T" "breakAfter"
            set_tcp(p[0.0,0.0,0.161,3.1415,0.0,0.0])
            movel(pose_trans(FRM_Reference, PSE_T), a=0.03, v=0.05)
          else:
            $ 1074 "Else" "noBreak"
            $ 1075 "'If random pose is out of reach, set the initial cam pose'"
            # 'If random pose is out of reach, set the initial cam pose'
            $ 1076 "PSE_T≔CAM_Pose"
            global PSE_T=CAM_Pose
            $ 1077 "PSE_T" "breakAfter"
            set_tcp(p[0.0,0.0,0.161,3.1415,0.0,0.0])
            movel(pose_trans(FRM_Reference, PSE_T), a=0.03, v=0.05)
          end
        end
        $ 1078 "Wait: 0.5"
        sleep(0.5)
        $ 1079 "Set"
        set_tcp(p[0.0,0.0,0.161,3.1415,0.0,0.0])
        # begin: URCap Program Node
        #   Source: SensoPart VISOR Robotic, 2.0.0, SensoPart Industriesensorik GmbH
        #   Type: VISOR Trigger
        $ 1080 "# 1 VISOR Trigger"
        visor_changeJob(1, "Object Detection Single", 6000)
        visor_trigger(1, 6000, "arm")
        # end: URCap Program Node
        $ 1081 "If visor_isResponseOk(1)"
        if ( visor_isResponseOk (1)):
          $ 1082 "CAM_CNT_Obj≔visor_partsFound(1)"
          global CAM_CNT_Obj= visor_partsFound (1)
          $ 1083 "CAM_OBJ_Pose≔visor_getPose3d(1, 0)"
          global CAM_OBJ_Pose= visor_getPose3d (1, 0)
          $ 1084 "If CAM_CNT_Obj>0"
          if (CAM_CNT_Obj>0):
            $ 1085 "CAM_OBJ_Color≔visor_getAdditionalData(1, 0)"
            global CAM_OBJ_Color= visor_getAdditionalData (1, 0)
            $ 1086 "CAM_DetectScore≔to_num(visor_getAdditionalData(1, 1))/1000"
            global CAM_DetectScore=to_num( visor_getAdditionalData (1, 1))/1000
            $ 1087 "OBJ_Detected≔ True "
            global OBJ_Detected=  True
          end
        else:
          $ 1088 "Else" "noBreak"
          $ 1089 "CAM_Captures≔CAM_Captures+1"
          global CAM_Captures=CAM_Captures+1
        end
        $ 1090 "If OBJ_Detected"
        if (OBJ_Detected):
          $ 1091 "Get object data"
          $ 1092 "PRC_CntDetect≔0"
          global PRC_CntDetect=0
          $ 1093 "Loop PRC_CntDetect<CAM_CNT_Obj"
          while (PRC_CntDetect<CAM_CNT_Obj):
            $ 1094 "get object and jig number"
            $ 1095 "If ITM_ID≟1 and JIG≟7"
            if (ITM_ID == 1  and  JIG == 7):
              $ 1096 "FRM_Reference≔FRM_Cap_SSRack"
              global FRM_Reference=FRM_Cap_SSRack
            else:
              $ 1097 "ElseIf ITM_ID≟5 and JIG≟7"
              if (ITM_ID == 5  and  JIG == 7):
                $ 1098 "FRM_Reference≔uLM_Cap_SSRack"
                global FRM_Reference=uLM_Cap_SSRack
              end
            end
            $ 1101 "PSE_T≔pose_trans(pose_inv(FRM_Reference), CAM_OBJ_Pose)"
            global PSE_T= pose_trans ( pose_inv (FRM_Reference), CAM_OBJ_Pose)
            $ 1102 "CAM_Result.append(get_pattern_counter(PSE_T, 'X', pattern=[10, 5], patternsize=[0.181, 0.081]))"
            CAM_Result.append(get_pattern_counter(PSE_T, "X", pattern=[10, 5], patternsize=[0.181, 0.081]))
            $ 1103 "PRC_CntDetect≔PRC_CntDetect+1"
            global PRC_CntDetect=PRC_CntDetect+1
          end
          $ 1104 "CAM_Done≔ True "
          global CAM_Done=  True
        else:
          $ 1105 "ElseIf CAM_Captures≥CAM_PRM_Retries"
          if (CAM_Captures >= CAM_PRM_Retries):
            $ 1106 "CAM_Done≔ True "
            global CAM_Done=  True
          else:
            $ 1107 "Else" "noBreak"
            $ 1108 "CAM_Captures≔CAM_Captures+1"
            global CAM_Captures=CAM_Captures+1
          end
        end
      end
    end
    $ 1109 "'=========='"
    # '=========='
    $ 1110 "PostSettings"
    $ 1111 "FRM_Reference≔p[0,0,0,0,0,0]"
    global FRM_Reference=p[0,0,0,0,0,0]
    $ 1112 "Set"
    set_tcp(p[0.0,0.0,0.161,3.1415,0.0,0.0])
    $ 1113 "CAM_Pose≔p[0,0,0,0,0,0]"
    global CAM_Pose=p[0,0,0,0,0,0]
    $ 1114 "Action≔0"
    global Action=0
    $ 1115 "Action_Info≔''"
    global Action_Info=""
  end
  def Sub_AMR_MiR_V3():
    $ 1116 "Sub_AMR_MiR_V3" "noBreak"
    $ 1117 "PreSettings"
    $ 1118 "AMR_TargetList≔[1,2,3,4,5,21,22,23,24,31,32,33,34,35,36,37,38,41]"
    global AMR_TargetList=[1,2,3,4,5,21,22,23,24,31,32,33,34,35,36,37,38,41]
    $ 1119 "AMR_Done≔ False "
    global AMR_Done=  False
    $ 1120 "AMR_PosActual≔T2O_Current_Pos"
    global AMR_PosActual=modbus_get_signal_status("T2O_Current_Pos")
    $ 1121 "AMR_Attemps≔T2O_Nav_Attemps"
    global AMR_Attemps=modbus_get_signal_status("T2O_Nav_Attemps")
    $ 1122 "AMR_Battery≔MiR_Battery_Lvl"
    global AMR_Battery=modbus_get_signal_status("MiR_Battery_Lvl")
    $ 1123 "AMR_Charging≔(T2O_Charging≟1)"
    global AMR_Charging=(modbus_get_signal_status("T2O_Charging") == 1)
    $ 1124 "AMR_Position≔struct(position_identifier=T2O_Current_Pos, x1=MiR_Position_X1, x2=MiR_Position_X2, y1=MiR_Position_Y1, y2=MiR_Position_Y2, theta1=MiR_Theta_1, theta2=MiR_Theta_2) "
    global AMR_Position=struct(position_identifier=modbus_get_signal_status("T2O_Current_Pos"), x1=modbus_get_signal_status("MiR_Position_X1"), x2=modbus_get_signal_status("MiR_Position_X2"), y1=modbus_get_signal_status("MiR_Position_Y1"), y2=modbus_get_signal_status("MiR_Position_Y2"), theta1=modbus_get_signal_status("MiR_Theta_1"), theta2=modbus_get_signal_status("MiR_Theta_2"))
    $ 1125 "If MiR_Mode≠7"
    if (modbus_get_signal_status("MiR_Mode") != 7):
      $ 1126 "Error"
      $ 1127 "set_error(ERROR_AMR_WRONG_MODE)"
      set_error(ERROR_AMR_WRONG_MODE)
      $ 1128 "AMR_Done≔ True "
      global AMR_Done=  True
    end
    $ 1129 "'=========='"
    # '=========='
    $ 1130 "Switch STATE"
    switch_1 = STATE
    $ 1131 "Case 1"
    if (1 == switch_1):
      $ 1132 "stopping"
      $ 1133 "If T2O_Done≟1 and O2T_Acknowledge≟0"
      if (modbus_get_signal_status("T2O_Done") == 1  and  modbus_get_signal_status("O2T_Acknowledge") == 0):
        $ 1134 "Set O2T_Acknowledge=1"
        modbus_set_output_register("O2T_Acknowledge", 1)
      end
      $ 1135 "Set MiR_CMD_Stop=On"
      modbus_set_output_signal("MiR_CMD_Stop", True)
      $ 1136 "AMR_Position.position_identifier = 0"
      AMR_Position.position_identifier = 0
      $ 1137 "AMR_Done≔ True "
      global AMR_Done=  True
    elif (2 == switch_1):
      $ 1138 "Case 2"
      $ 1139 "stopped"
      $ 1140 "If MiR_State≠3 and MiR_State≠5"
      if (modbus_get_signal_status("MiR_State") != 3  and  modbus_get_signal_status("MiR_State") != 5):
        $ 1141 "Set MiR_CMD_Stop=Off"
        modbus_set_output_signal("MiR_CMD_Stop", False)
      end
    elif (3 == switch_1):
      $ 1142 "Case 3"
      $ 1143 "resetting"
      $ 1144 "Set O2T_Mis_Main=Off"
      modbus_set_output_signal("O2T_Mis_Main", False)
      $ 1145 "Set O2T_Mis_Charge=Off"
      modbus_set_output_signal("O2T_Mis_Charge", False)
      $ 1146 "If MiR_Mis_Queue>0"
      if (modbus_get_signal_status("MiR_Mis_Queue")>0):
        $ 1147 "Set MiR_CMD_Clear_Q=On"
        modbus_set_output_signal("MiR_CMD_Clear_Q", True)
        $ 1148 "Wait MiR_Mis_Queue≟0"
        while (not(modbus_get_signal_status("MiR_Mis_Queue") == 0)):
          sync()
        end
        $ 1149 "Set MiR_CMD_Clear_Q=Off"
        modbus_set_output_signal("MiR_CMD_Clear_Q", False)
      end
      $ 1150 "If MiR_Error_ID≠0"
      if (modbus_get_signal_status("MiR_Error_ID") != 0):
        $ 1151 "Set MiR_CMD_Clear_E=On"
        modbus_set_output_signal("MiR_CMD_Clear_E", True)
        $ 1152 "Wait MiR_Error_ID≟0"
        while (not(modbus_get_signal_status("MiR_Error_ID") == 0)):
          sync()
        end
        $ 1153 "Set MiR_CMD_Clear_E=Off"
        modbus_set_output_signal("MiR_CMD_Clear_E", False)
      end
      $ 1154 "Set O2T_Action=0"
      modbus_set_output_register("O2T_Action", 0)
      $ 1155 "Set O2T_Acknowledge=0"
      modbus_set_output_register("O2T_Acknowledge", 0)
      $ 1156 "Set O2T_Target_Pos=0"
      modbus_set_output_register("O2T_Target_Pos", 0)
      $ 1157 "Set O2T_Footprint=0"
      modbus_set_output_register("O2T_Footprint", 0)
      $ 1158 "Set O2T_ProtectOff=0"
      modbus_set_output_register("O2T_ProtectOff", 0)
      $ 1159 "Set O2T_Dock=0"
      modbus_set_output_register("O2T_Dock", 0)
      $ 1160 "AMR_Attemps≔0"
      global AMR_Attemps=0
      $ 1161 "AMR_PosTarget≔0"
      global AMR_PosTarget=0
      $ 1162 "AMR_Step≔0"
      global AMR_Step=0
      $ 1163 "AMR_AtTarget≔ False "
      global AMR_AtTarget=  False
      $ 1164 "If MiR_State≟4 or MiR_State≟3 or MiR_State≟10"
      if (modbus_get_signal_status("MiR_State") == 4  or  modbus_get_signal_status("MiR_State") == 3  or  modbus_get_signal_status("MiR_State") == 10):
        $ 1165 "AMR_Done≔ True "
        global AMR_Done=  True
      end
    elif (5 == switch_1):
      $ 1166 "Case 5"
      $ 1167 "starting"
      $ 1168 "If MiR_State≟4"
      if (modbus_get_signal_status("MiR_State") == 4):
        $ 1169 "Set MiR_CMD_Start=On"
        modbus_set_output_signal("MiR_CMD_Start", True)
        $ 1170 "Wait MiR_State≠4"
        while (not(modbus_get_signal_status("MiR_State") != 4)):
          sync()
        end
        $ 1171 "Set MiR_CMD_Start=Off"
        modbus_set_output_signal("MiR_CMD_Start", False)
        $ 1172 "AMR_Done≔ True "
        global AMR_Done=  True
      else:
        $ 1173 "ElseIf MiR_State≟10"
        if (modbus_get_signal_status("MiR_State") == 10):
          $ 1174 "'MiR in protective stop. Wait'"
          # 'MiR in protective stop. Wait'
          $ 1175 "AMR_Done≔ True "
          global AMR_Done=  True
        else:
          $ 1176 "ElseIf MiR_State≟3"
          if (modbus_get_signal_status("MiR_State") == 3):
            $ 1177 "AMR_Done≔ True "
            global AMR_Done=  True
          end
        end
      end
    elif (6 == switch_1):
      $ 1178 "Case 6"
      $ 1179 "execute"
      $ 1180 "AMR_AtTarget≔(AMR_PosActual≟AMR_PosTarget)"
      global AMR_AtTarget=(AMR_PosActual == AMR_PosTarget)
      $ 1181 "Switch AMR_Step"
      switch_2 = AMR_Step
      $ 1182 "Case 0"
      if (0 == switch_2):
        $ 1183 "If  not AMR_AtTarget"
        if (  not  AMR_AtTarget):
          $ 1184 "AMR_Step≔1"
          global AMR_Step=1
        else:
          $ 1185 "Else" "noBreak"
          $ 1186 "AMR_Done≔ True "
          global AMR_Done=  True
        end
      elif (1 == switch_2):
        $ 1187 "Case 1"
        $ 1188 "general Settings"
        $ 1189 "Set O2T_Acknowledge=0"
        modbus_set_output_register("O2T_Acknowledge", 0)
        $ 1190 "check for error"
        $ 1191 "If OBJ_Picked and MiR_State≟10"
        if (OBJ_Picked  and  modbus_get_signal_status("MiR_State") == 10):
          $ 1192 "Error"
          $ 1193 "set_error(ERROR_ROBOT_ARM_NOT_IN_HOME_POSE)"
          set_error(ERROR_ROBOT_ARM_NOT_IN_HOME_POSE)
          $ 1194 "Action≔0"
          global Action=0
        else:
          $ 1195 "ElseIf  not found_in_list(AMR_PosTarget, AMR_TargetList)"
          if (  not  found_in_list(AMR_PosTarget, AMR_TargetList)):
            $ 1196 "Error"
            $ 1197 "set_error(ERROR_UNKNOWN_POSE)"
            set_error(ERROR_UNKNOWN_POSE)
            $ 1198 "Action≔0"
            global Action=0
          end
        end
        $ 1199 "If MiR_State≟3"
        if (modbus_get_signal_status("MiR_State") == 3):
          $ 1200 "Set MiR_CMD_Start=Off"
          modbus_set_output_signal("MiR_CMD_Start", False)
          $ 1201 "Switch Action"
          switch_3 = Action
          $ 1202 "Case 51"
          if (51 == switch_3):
            $ 1203 "Charge"
            $ 1204 "'trigger the charging mission'"
            # 'trigger the charging mission'
            $ 1205 "'target pos is predefined'"
            # 'target pos is predefined'
            $ 1206 "Set O2T_Footprint=0"
            modbus_set_output_register("O2T_Footprint", 0)
            $ 1207 "Set O2T_Action=1"
            modbus_set_output_register("O2T_Action", 1)
            $ 1208 "If MiR_Mis_Queue≟0"
            if (modbus_get_signal_status("MiR_Mis_Queue") == 0):
              $ 1209 "Set O2T_Mis_Charge=On"
              modbus_set_output_signal("O2T_Mis_Charge", True)
              $ 1210 "Wait MiR_Mis_Queue≥1"
              while (not(modbus_get_signal_status("MiR_Mis_Queue") >= 1)):
                sync()
              end
              $ 1211 "Set O2T_Mis_Charge=Off"
              modbus_set_output_signal("O2T_Mis_Charge", False)
            end
          elif (52 == switch_3):
            $ 1212 "Case 52"
            $ 1213 "Navigate"
            $ 1214 "'trigger the standard missoin'"
            # 'trigger the standard missoin'
            $ 1215 "Set O2T_Footprint=AMR_FootprintID"
            modbus_set_output_register("O2T_Footprint", AMR_FootprintID)
            $ 1216 "Set O2T_Target_Pos=AMR_PosTarget"
            modbus_set_output_register("O2T_Target_Pos", AMR_PosTarget)
            $ 1217 "Set O2T_Action=2"
            modbus_set_output_register("O2T_Action", 2)
            $ 1218 "If MiR_Mis_Queue≟0"
            if (modbus_get_signal_status("MiR_Mis_Queue") == 0):
              $ 1219 "Set O2T_Mis_Main=On"
              modbus_set_output_signal("O2T_Mis_Main", True)
              $ 1220 "Wait MiR_Mis_Queue≥1"
              while (not(modbus_get_signal_status("MiR_Mis_Queue") >= 1)):
                sync()
              end
              $ 1221 "Set O2T_Mis_Main=Off"
              modbus_set_output_signal("O2T_Mis_Main", False)
            end
          end
        else:
          $ 1222 "ElseIf MiR_State≟4"
          if (modbus_get_signal_status("MiR_State") == 4):
            $ 1223 "Set MiR_CMD_Start=On"
            modbus_set_output_signal("MiR_CMD_Start", True)
          else:
            $ 1224 "ElseIf MiR_State≟5"
            if (modbus_get_signal_status("MiR_State") == 5):
              $ 1225 "AMR_Step≔2"
              global AMR_Step=2
            else:
              $ 1226 "ElseIf MiR_State≟10"
              if (modbus_get_signal_status("MiR_State") == 10):
                $ 1227 "'AMR still in safeguard stop'"
                # 'AMR still in safeguard stop'
              end
            end
          end
        end
      elif (2 == switch_2):
        $ 1228 "Case 2"
        $ 1229 "acknowledge handshake"
        $ 1230 "If T2O_Done≟1 and O2T_Acknowledge≟0"
        if (modbus_get_signal_status("T2O_Done") == 1  and  modbus_get_signal_status("O2T_Acknowledge") == 0):
          $ 1231 "Set O2T_Acknowledge=1"
          modbus_set_output_register("O2T_Acknowledge", 1)
        else:
          $ 1232 "ElseIf T2O_Done≟0 and O2T_Acknowledge≟1"
          if (modbus_get_signal_status("T2O_Done") == 0  and  modbus_get_signal_status("O2T_Acknowledge") == 1):
            $ 1233 "Set O2T_Acknowledge=0"
            modbus_set_output_register("O2T_Acknowledge", 0)
            $ 1234 "AMR_AtTarget≔(AMR_PosActual≟AMR_PosTarget)"
            global AMR_AtTarget=(AMR_PosActual == AMR_PosTarget)
            $ 1235 "AMR_Done≔ True "
            global AMR_Done=  True
          end
        end
      end
      $ 1236 "translate errors"
      $ 1237 "If AMR_Done"
      if (AMR_Done):
        $ 1238 "Switch T2O_Error_ID"
        switch_2 = modbus_get_signal_status("T2O_Error_ID")
        $ 1239 "Case 2003"
        if (2003 == switch_2):
          $ 1240 "error"
          $ 1241 "set_error(ERROR_NOT_DOCKED)"
          set_error(ERROR_NOT_DOCKED)
        elif (2007 == switch_2):
          $ 1242 "Case 2007"
          $ 1243 "error"
          $ 1244 "set_error(ERROR_NOT_REACHABLE_TARGET)"
          set_error(ERROR_NOT_REACHABLE_TARGET)
        elif (2008 == switch_2):
          $ 1245 "Case 2008"
          $ 1246 "error"
          $ 1247 "set_error(ERROR_CHARGING_NOT_STARTED)"
          set_error(ERROR_CHARGING_NOT_STARTED)
        end
      end
    elif (7 == switch_1):
      $ 1248 "Case 7"
      $ 1249 "completing"
      $ 1250 "If MiR_Mis_Queue>0"
      if (modbus_get_signal_status("MiR_Mis_Queue")>0):
        $ 1251 "Set MiR_CMD_Abort=On"
        modbus_set_output_signal("MiR_CMD_Abort", True)
        $ 1252 "Wait MiR_Mis_Queue≟0"
        while (not(modbus_get_signal_status("MiR_Mis_Queue") == 0)):
          sync()
        end
        $ 1253 "Set MiR_CMD_Abort=Off"
        modbus_set_output_signal("MiR_CMD_Abort", False)
      end
      $ 1254 "If MiR_State≟3 or MiR_State≟10"
      if (modbus_get_signal_status("MiR_State") == 3  or  modbus_get_signal_status("MiR_State") == 10):
        $ 1255 "AMR_Done≔ True "
        global AMR_Done=  True
      end
    elif (9 == switch_1):
      $ 1256 "Case 9"
      $ 1257 "holding"
      $ 1258 "Set MiR_CMD_Abort=On"
      modbus_set_output_signal("MiR_CMD_Abort", True)
      $ 1259 "If MiR_State≟3 or MiR_State≟10"
      if (modbus_get_signal_status("MiR_State") == 3  or  modbus_get_signal_status("MiR_State") == 10):
        $ 1260 "Set MiR_CMD_Abort=Off"
        modbus_set_output_signal("MiR_CMD_Abort", False)
        $ 1261 "AMR_Done≔ True "
        global AMR_Done=  True
      end
    elif (11 == switch_1):
      $ 1262 "Case 11"
      $ 1263 "unholding"
      $ 1264 "Set MiR_CMD_Start=On"
      modbus_set_output_signal("MiR_CMD_Start", True)
      $ 1265 "If MiR_State≠4"
      if (modbus_get_signal_status("MiR_State") != 4):
        $ 1266 "Set MiR_CMD_Start=Off"
        modbus_set_output_signal("MiR_CMD_Start", False)
        $ 1267 "AMR_Step≔0"
        global AMR_Step=0
        $ 1268 "AMR_Done≔ True "
        global AMR_Done=  True
      end
    elif (12 == switch_1):
      $ 1269 "Case 12"
      $ 1270 "suspending"
      $ 1271 "'none'"
      # 'none'
    elif (14 == switch_1):
      $ 1272 "Case 14"
      $ 1273 "unsuspending"
      $ 1274 "'none'"
      # 'none'
    elif (15 == switch_1):
      $ 1275 "Case 15"
      $ 1276 "aborting"
      $ 1277 "Set MiR_CMD_Abort=On"
      modbus_set_output_signal("MiR_CMD_Abort", True)
      $ 1278 "Wait MiR_State≟3"
      while (not(modbus_get_signal_status("MiR_State") == 3)):
        sync()
      end
      $ 1279 "Set MiR_CMD_Abort=Off"
      modbus_set_output_signal("MiR_CMD_Abort", False)
    elif (17 == switch_1):
      $ 1280 "Case 17"
      $ 1281 "clearing"
      $ 1282 "If MiR_Error_ID≠0"
      if (modbus_get_signal_status("MiR_Error_ID") != 0):
        $ 1283 "Set MiR_CMD_Clear_E=On"
        modbus_set_output_signal("MiR_CMD_Clear_E", True)
        $ 1284 "Wait MiR_Error_ID≟0"
        while (not(modbus_get_signal_status("MiR_Error_ID") == 0)):
          sync()
        end
        $ 1285 "Set MiR_CMD_Clear_E=Off"
        modbus_set_output_signal("MiR_CMD_Clear_E", False)
      end
      $ 1286 "If MiR_Error_ID≟0"
      if (modbus_get_signal_status("MiR_Error_ID") == 0):
        $ 1287 "AMR_Done≔ True "
        global AMR_Done=  True
      end
    end
    $ 1288 "'=========='"
    # '=========='
    $ 1289 "PostSettings"
    $ 1290 "AMR_Position≔struct(position_identifier=T2O_Current_Pos, x1=MiR_Position_X1, x2=MiR_Position_X2, y1=MiR_Position_Y1, y2=MiR_Position_Y2, theta1=MiR_Theta_1, theta2=MiR_Theta_2) "
    global AMR_Position=struct(position_identifier=modbus_get_signal_status("T2O_Current_Pos"), x1=modbus_get_signal_status("MiR_Position_X1"), x2=modbus_get_signal_status("MiR_Position_X2"), y1=modbus_get_signal_status("MiR_Position_Y1"), y2=modbus_get_signal_status("MiR_Position_Y2"), theta1=modbus_get_signal_status("MiR_Theta_1"), theta2=modbus_get_signal_status("MiR_Theta_2"))
  end
  def Sub_Action_V4():
    $ 1291 "Sub_Action_V4" "noBreak"
    $ 1292 "PreSettings"
    $ 1293 "init poses"
    $ 1294 "PSE_A≔p[0,0,0,0,0,0]"
    global PSE_A=p[0,0,0,0,0,0]
    $ 1295 "PSE_A_H≔p[0,0,0,0,0,0]"
    global PSE_A_H=p[0,0,0,0,0,0]
    $ 1296 "PSE_T≔p[0,0,0,0,0,0]"
    global PSE_T=p[0,0,0,0,0,0]
    $ 1297 "PSE_T_H≔p[0,0,0,0,0,0]"
    global PSE_T_H=p[0,0,0,0,0,0]
    $ 1298 "PSE_G≔p[0,0,0,0,0,0]"
    global PSE_G=p[0,0,0,0,0,0]
    $ 1299 "PSE_G_H≔p[0,0,0,0,0,0]"
    global PSE_G_H=p[0,0,0,0,0,0]
    $ 1300 "PSE_R≔p[0,0,0,0,0,0]"
    global PSE_R=p[0,0,0,0,0,0]
    $ 1301 "PSE_R_H≔p[0,0,0,0,0,0]"
    global PSE_R_H=p[0,0,0,0,0,0]
    $ 1302 "JNT_Q≔[0,0,0,0,0,0]"
    global JNT_Q=[0,0,0,0,0,0]
    $ 1303 "JNT_S≔[0,0,0,0,0,0]"
    global JNT_S=[0,0,0,0,0,0]
    $ 1304 "Gripping parameters"
    $ 1305 "OBJ = find_object_by_type(OBJs, OBJ_Type)"
    OBJ = find_object_by_type(OBJs, OBJ_Type)
    $ 1306 "GRP_Open_Pos≔OBJ.dimension.diameter * 1000 + 6"
    global GRP_Open_Pos=OBJ.dimension.diameter * 1000 + 6
    $ 1307 "GRP_Offset≔OBJ.gripper_offset"
    global GRP_Offset=OBJ.gripper_offset
    $ 1308 "rq_set_force_norm(50)"
     rq_set_force_norm (50)
    $ 1309 "rq_set_speed_norm(50)"
     rq_set_speed_norm (50)
    $ 1310 "Switch ITM_ID"
    switch_1 = ITM_ID
    $ 1311 "Case 1"
    if (1 == switch_1):
      $ 1312 "uML"
      $ 1313 "JIG2 = find_object_by_type(JIGs, JIG)"
      JIG2 = find_object_by_type(JIGs, JIG)
      $ 1314 "JIG_Offset≔JIG2.jig_offset"
      global JIG_Offset=JIG2.jig_offset
      $ 1315 "Switch JIG"
      switch_2 = JIG
      $ 1316 "Case 1"
      if (1 == switch_2):
        $ 1317 "3FG"
        $ 1318 "define poses"
        $ 1319 "FRM_Reference≔ULM_3FG"
        global FRM_Reference=ULM_3FG
        $ 1320 "JNT_Q≔JNT_HOME"
        global JNT_Q=JNT_HOME
        $ 1321 "PSE_T≔pose_trans(GRP_Offset, JIG_Offset)"
        global PSE_T= pose_trans (GRP_Offset, JIG_Offset)
        $ 1322 "PSE_A≔pose_trans(PSE_T, p[0,0,0.100,0,0,0])"
        global PSE_A= pose_trans (PSE_T, p[0,0,0.100,0,0,0])
        $ 1323 "PSE_R≔pose_add(PSE_T, p[0,0,0.100,0,0,0])"
        global PSE_R= pose_add (PSE_T, p[0,0,0.100,0,0,0])
      elif (2 == switch_2):
        $ 1324 "Case 2"
        $ 1325 "Input"
        $ 1326 "'CHANGE THE REFERENCE TO THE FRAME TO MOVE IN'"
        # 'CHANGE THE REFERENCE TO THE FRAME TO MOVE IN'
        $ 1327 "define poses"
        $ 1328 "FRM_Reference≔ULM_Input"
        global FRM_Reference=ULM_Input
        $ 1329 "PSE_T≔pose_trans(pose_trans(get_pattern_pos_rectangle(OBJ_Nbr, 'X', [10,5], patternsize=[0.181,0.081]), GRP_Offset), JIG_Offset)"
        global PSE_T= pose_trans ( pose_trans (get_pattern_pos_rectangle(OBJ_Nbr, "X", [10,5], patternsize=[0.181,0.081]), GRP_Offset), JIG_Offset)
        $ 1330 "If Action≟1"
        if (Action == 1):
          $ 1331 "PSE_R≔pose_add(PSE_T, p[0,0,0.200,0,0,0])"
          global PSE_R= pose_add (PSE_T, p[0,0,0.200,0,0,0])
          $ 1332 "PSE_A≔pose_add(PSE_T, p[0,0,0.100,0,0,0])"
          global PSE_A= pose_add (PSE_T, p[0,0,0.100,0,0,0])
        else:
          $ 1333 "ElseIf Action≟2"
          if (Action == 2):
            $ 1334 "PSE_R≔pose_add(PSE_T, p[0,0,0.100,0,0,0])"
            global PSE_R= pose_add (PSE_T, p[0,0,0.100,0,0,0])
            $ 1335 "PSE_A≔pose_add(PSE_T, p[0,0,0.200,0,0,0])"
            global PSE_A= pose_add (PSE_T, p[0,0,0.200,0,0,0])
          end
        end
      elif (3 == switch_2):
        $ 1336 "Case 3"
        $ 1337 "Output"
        $ 1338 "'CHANGE THE REFERENCE TO THE FRAME TO MOVE IN'"
        # 'CHANGE THE REFERENCE TO THE FRAME TO MOVE IN'
        $ 1339 "define poses"
        $ 1340 "FRM_Reference≔ULM_Output"
        global FRM_Reference=ULM_Output
        $ 1341 "PSE_T≔pose_trans(pose_trans(get_pattern_pos_rectangle(OBJ_Nbr, 'X', [10,5], patternsize=[0.181,0.081]), GRP_Offset), JIG_Offset)"
        global PSE_T= pose_trans ( pose_trans (get_pattern_pos_rectangle(OBJ_Nbr, "X", [10,5], patternsize=[0.181,0.081]), GRP_Offset), JIG_Offset)
        $ 1343 "If Action≟1"
        if (Action == 1):
          $ 1344 "PSE_R≔pose_add(PSE_T, p[0,0,0.200,0,0,0])"
          global PSE_R= pose_add (PSE_T, p[0,0,0.200,0,0,0])
          $ 1345 "PSE_A≔pose_add(PSE_T, p[0,0,0.100,0,0,0])"
          global PSE_A= pose_add (PSE_T, p[0,0,0.100,0,0,0])
        else:
          $ 1346 "ElseIf Action≟2"
          if (Action == 2):
            $ 1347 "PSE_R≔pose_add(PSE_T, p[0,0,0.100,0,0,0])"
            global PSE_R= pose_add (PSE_T, p[0,0,0.100,0,0,0])
            $ 1348 "PSE_A≔pose_add(PSE_T, p[0,0,0.200,0,0,0])"
            global PSE_A= pose_add (PSE_T, p[0,0,0.200,0,0,0])
          end
        end
      elif (4 == switch_2):
        $ 1349 "Case 4"
        $ 1350 "jig centrifuge racks"
        $ 1351 "define poses"
        $ 1352 "FRM_Reference≔ULM_Cent_Racks"
        global FRM_Reference=ULM_Cent_Racks
        $ 1353 "PSE_T≔get_pattern_pos_rectangle(JIG_Slot, 'X', [4,1], patternsize=[0.291,0])"
        global PSE_T=get_pattern_pos_rectangle(JIG_Slot, "X", [4,1], patternsize=[0.291,0])
        $ 1354 "If OBJ_Nbr≠0"
        if (OBJ_Nbr != 0):
          $ 1355 "PSE_T≔pose_trans(pose_trans(PSE_T, get_pattern_pos_rectangle(OBJ_Nbr, 'X', [3,3], patternsize=[0.060,0.060])),p[-0.030, -0.030,0,0,0,3.927])"
          global PSE_T= pose_trans ( pose_trans (PSE_T, get_pattern_pos_rectangle(OBJ_Nbr, "X", [3,3], patternsize=[0.060,0.060])),p[-0.030, -0.030,0,0,0,3.927])
        end
        $ 1356 "PSE_T≔pose_trans(PSE_T, GRP_Offset)"
        global PSE_T= pose_trans (PSE_T, GRP_Offset)
        $ 1357 "If Action≟1"
        if (Action == 1):
          $ 1358 "PSE_R≔pose_add(PSE_T, p[0,0,0.200,0,0,0])"
          global PSE_R= pose_add (PSE_T, p[0,0,0.200,0,0,0])
          $ 1359 "PSE_A≔pose_add(PSE_T, p[0,0,0.100,0,0,0])"
          global PSE_A= pose_add (PSE_T, p[0,0,0.100,0,0,0])
        else:
          $ 1360 "ElseIf Action≟2"
          if (Action == 2):
            $ 1361 "PSE_R≔pose_add(PSE_T, p[0,0,0.100,0,0,0])"
            global PSE_R= pose_add (PSE_T, p[0,0,0.100,0,0,0])
            $ 1362 "PSE_A≔pose_add(PSE_T, p[0,0,0.200,0,0,0])"
            global PSE_A= pose_add (PSE_T, p[0,0,0.200,0,0,0])
          end
        end
      elif (6 == switch_2):
        $ 1363 "Case 6"
        $ 1364 "Caps bin"
        $ 1365 "define poses"
        $ 1366 "'Drop cap'"
        # 'Drop cap'
        $ 1367 "FRM_Reference=ULM_Cap_Bin"
        FRM_Reference=ULM_Cap_Bin
        $ 1368 "PSE_T≔pose_RPY2RotVec(p[0,0,0,0,0,0])"
        global PSE_T=pose_RPY2RotVec(p[0,0,0,0,0,0])
        $ 1369 "PSE_T_H≔pose_add(PSE_T, p[0,0,-0.011,0,0,0])"
        global PSE_T_H= pose_add (PSE_T, p[0,0,-0.011,0,0,0])
        $ 1370 "PSE_A≔pose_trans(PSE_T, p[0,0,0.1,0,0,0])"
        global PSE_A= pose_trans (PSE_T, p[0,0,0.1,0,0,0])
        $ 1371 "PSE_R_H≔pose_add(PSE_T, p[0,0,0.100,0,0,0])"
        global PSE_R_H= pose_add (PSE_T, p[0,0,0.100,0,0,0])
        $ 1372 "PSE_R≔pose_add(PSE_T, p[0,0,0.100,0,0,0])"
        global PSE_R= pose_add (PSE_T, p[0,0,0.100,0,0,0])
      elif (7 == switch_2):
        $ 1373 "Case 7"
        $ 1374 "Sarstedt"
        $ 1375 "'CHANGE THE REFERENCE TO THE FRAME TO MOVE IN'"
        # 'CHANGE THE REFERENCE TO THE FRAME TO MOVE IN'
        $ 1381 "If TASK.ID≟10"
        if (TASK.ID == 10):
          $ 1382 "Frame & Position Params"
          $ 1384 "FRM_Reference = CAM_LM_SSRack"
          FRM_Reference = CAM_LM_SSRack
          $ 1389 "PSE_T≔uLM_SS_PickPlc"
          global PSE_T=uLM_SS_PickPlc
          $ 1390 "PSE_A≔pose_trans(PSE_T, p[0,0,0.1,0,0,0])"
          global PSE_A= pose_trans (PSE_T, p[0,0,0.1,0,0,0])
          $ 1391 "PSE_R≔pose_add(PSE_T, p[0,0,0.1,0,0,0])"
          global PSE_R= pose_add (PSE_T, p[0,0,0.1,0,0,0])
        else:
          $ 1392 "ElseIf TASK.ID≟11"
          if (TASK.ID == 11):
            $ 1393 "FRM_Reference = ULM_SS_Jig"
            FRM_Reference = ULM_SS_Jig
            $ 1394 "PSE_T≔pose_RPY2RotVec(p[0,0,0,0,0,0])"
            global PSE_T=pose_RPY2RotVec(p[0,0,0,0,0,0])
            $ 1395 "PSE_T≔pose_trans(PSE_T, GRP_Offset)"
            global PSE_T=pose_trans(PSE_T, GRP_Offset)
            $ 1396 "PSE_A≔pose_trans(PSE_T, p[0,0,0.1,0,0,0])"
            global PSE_A= pose_trans (PSE_T, p[0,0,0.1,0,0,0])
            $ 1397 "PSE_R≔pose_add(PSE_T, p[0,0,0.2,0,0,0])"
            global PSE_R= pose_add (PSE_T, p[0,0,0.2,0,0,0])
          end
        end
      elif (8 == switch_2):
        $ 1398 "Case 8"
        $ 1399 "NoK"
        $ 1400 "define poses"
        $ 1401 "'NoK'"
        # 'NoK'
        $ 1402 "FRM_Reference=ULM_NoK"
        FRM_Reference=ULM_NoK
        $ 1403 "PSE_T≔pose_RPY2RotVec(p[0,0,0,0,0,0])"
        global PSE_T=pose_RPY2RotVec(p[0,0,0,0,0,0])
        $ 1404 "PSE_A≔pose_trans(PSE_T, p[0,0,0.1,0,0,0])"
        global PSE_A= pose_trans (PSE_T, p[0,0,0.1,0,0,0])
        $ 1405 "PSE_R≔pose_add(PSE_T, p[0,0,0.100,0,0,0])"
        global PSE_R= pose_add (PSE_T, p[0,0,0.100,0,0,0])
      elif (9 == switch_2):
        $ 1406 "Case 9"
        $ 1407 "Pick_bott_jig"
        $ 1408 "define poses"
        $ 1409 "'NoK'"
        # 'NoK'
        $ 1410 "FRM_Reference=ULM_bottle_pick_const"
        FRM_Reference=p[0.08175869478771049,-0.47602162643540935,0.09,0.00141829700319658,-0.0027789445191063835,0.07763675748118615]
        $ 1411 "PSE_T≔pose_RPY2RotVec(p[0,0,0,0,0,0])"
        global PSE_T=pose_RPY2RotVec(p[0,0,0,0,0,0])
        $ 1412 "PSE_A≔pose_trans(PSE_T, p[0,0,0.1,0,0,0])"
        global PSE_A= pose_trans (PSE_T, p[0,0,0.1,0,0,0])
        $ 1413 "PSE_R≔pose_add(PSE_T, p[0,0,0.100,0,0,0])"
        global PSE_R= pose_add (PSE_T, p[0,0,0.100,0,0,0])
      elif (10 == switch_2):
        $ 1414 "Case 10"
        $ 1415 "Place_bott_jig"
        $ 1416 "define poses"
        $ 1417 "'NoK'"
        # 'NoK'
        $ 1418 "FRM_Reference=ULM_bottle_plac_const"
        FRM_Reference=p[-0.09502738395762109,-0.5154087721098056,0.095,0.0014590126708889871,-0.0028280855286173575,0.07763149296298452]
        $ 1419 "PSE_T≔pose_RPY2RotVec(p[0,0,0,0,0,0])"
        global PSE_T=pose_RPY2RotVec(p[0,0,0,0,0,0])
        $ 1420 "PSE_A≔pose_trans(PSE_T, p[0,0,0.1,0,0,0])"
        global PSE_A= pose_trans (PSE_T, p[0,0,0.1,0,0,0])
        $ 1421 "PSE_R≔pose_add(PSE_T, p[0,0,0.100,0,0,0])"
        global PSE_R= pose_add (PSE_T, p[0,0,0.100,0,0,0])
      elif (11 == switch_2):
        $ 1422 "Case 11"
        $ 1423 "Place_bott_jig"
        $ 1424 "define poses"
        $ 1425 "'NoK'"
        # 'NoK'
        $ 1426 "FRM_Reference=shake"
        FRM_Reference=shake
        $ 1427 "PSE_T≔pose_RPY2RotVec(p[0,0,0,0,0,0])"
        global PSE_T=pose_RPY2RotVec(p[0,0,0,0,0,0])
        $ 1428 "PSE_A≔pose_trans(PSE_T, p[0,0,0,0,0,0])"
        global PSE_A= pose_trans (PSE_T, p[0,0,0,0,0,0])
        $ 1429 "PSE_R≔pose_add(PSE_T, p[0,0,0,0,0,0])"
        global PSE_R= pose_add (PSE_T, p[0,0,0,0,0,0])
      elif (12 == switch_2):
        $ 1430 "Case 12"
        $ 1431 "Pick_Vial_jig"
        $ 1432 "define poses"
        $ 1433 "'NoK'"
        # 'NoK'
        $ 1434 "FRM_Reference=shake"
        FRM_Reference=shake
        $ 1435 "PSE_T≔pose_RPY2RotVec(p[0,0,0,0,0,0])"
        global PSE_T=pose_RPY2RotVec(p[0,0,0,0,0,0])
        $ 1436 "PSE_A≔pose_trans(PSE_T, p[0,0,0,0,0,0])"
        global PSE_A= pose_trans (PSE_T, p[0,0,0,0,0,0])
        $ 1437 "PSE_R≔pose_add(PSE_T, p[0,0,0,0,0,0])"
        global PSE_R= pose_add (PSE_T, p[0,0,0,0,0,0])
      end
    elif (2 == switch_1):
      $ 1438 "Case 2"
      $ 1439 "Centrifuge"
      $ 1440 "'CHANGE THE REFERENCE TO THE FRAME TO MOVE IN'"
      # 'CHANGE THE REFERENCE TO THE FRAME TO MOVE IN'
      $ 1441 "define poses"
      $ 1442 "FRM_Reference≔FRM_Centrifuge"
      global FRM_Reference=FRM_Centrifuge
      $ 1443 "PSE_T≔GRP_Offset"
      global PSE_T=GRP_Offset
      $ 1444 "If Action≟8"
      if (Action == 8):
        $ 1445 "PSE_R≔pose_add(PSE_T, p[0,0,0.250,0,0,0])"
        global PSE_R= pose_add (PSE_T, p[0,0,0.250,0,0,0])
        $ 1446 "PSE_A≔pose_add(PSE_T, p[0,0,0.150,0,0,0])"
        global PSE_A= pose_add (PSE_T, p[0,0,0.150,0,0,0])
      else:
        $ 1447 "ElseIf Action≟7"
        if (Action == 7):
          $ 1448 "PSE_R≔pose_add(PSE_T, p[0,0,0.150,0,0,0])"
          global PSE_R= pose_add (PSE_T, p[0,0,0.150,0,0,0])
          $ 1449 "PSE_A≔pose_add(PSE_T, p[0,0,0.250,0,0,0])"
          global PSE_A= pose_add (PSE_T, p[0,0,0.250,0,0,0])
        end
      end
    elif (3 == switch_1):
      $ 1450 "Case 3"
      $ 1451 "Output"
      $ 1452 "'CHANGE THE REFERENCE TO THE FRAME TO MOVE IN'"
      # 'CHANGE THE REFERENCE TO THE FRAME TO MOVE IN'
      $ 1453 "define poses"
      $ 1454 "FRM_Reference≔Base_const"
      global FRM_Reference=p[0.0,0.0,0.0,0.0,0.0,0.0]
      $ 1455 "PSE_T≔p[0,0,0,0,0,0]"
      global PSE_T=p[0,0,0,0,0,0]
      $ 1456 "PSE_A≔pose_add(PSE_T, p[0,0,0.150,0,0,0])"
      global PSE_A= pose_add (PSE_T, p[0,0,0.150,0,0,0])
      $ 1457 "PSE_R≔pose_add(PSE_T, p[0,0,0.100,0,0,0])"
      global PSE_R= pose_add (PSE_T, p[0,0,0.100,0,0,0])
    elif (5 == switch_1):
      $ 1458 "Case 5"
      $ 1459 "Sarstedt Pickup Table"
      $ 1460 "'CHANGE THE REFERENCE TO THE FRAME TO MOVE IN'"
      # 'CHANGE THE REFERENCE TO THE FRAME TO MOVE IN'
      $ 1461 "Switch JIG"
      switch_2 = JIG
      $ 1462 "Case 7"
      if (7 == switch_2):
        $ 1475 "Sarstedt"
        $ 1476 "'CHANGE THE REFERENCE TO THE FRAME TO MOVE IN'"
        # 'CHANGE THE REFERENCE TO THE FRAME TO MOVE IN'
        $ 1482 "If TASK.ID≟10"
        if (TASK.ID == 10):
          $ 1483 "Frame & Position Params"
          $ 1484 "FRM_Reference = CAM_LM_SSRack"
          FRM_Reference = CAM_LM_SSRack
          $ 1485 "PSE_T≔uLM_SS_PickPlc"
          global PSE_T=uLM_SS_PickPlc
          $ 1486 "PSE_A≔pose_trans(PSE_T, p[0,0,0.1,0,0,0])"
          global PSE_A= pose_trans (PSE_T, p[0,0,0.1,0,0,0])
          $ 1487 "PSE_R≔pose_add(PSE_T, p[0,0,0.1,0,0,0])"
          global PSE_R= pose_add (PSE_T, p[0,0,0.1,0,0,0])
        end
      end
    elif (13 == switch_1):
      $ 1494 "Case 13"
      $ 1495 "Sarstedt Pickup Table"
      $ 1496 "'CHANGE THE REFERENCE TO THE FRAME TO MOVE IN'"
      # 'CHANGE THE REFERENCE TO THE FRAME TO MOVE IN'
      $ 1497 "Switch JIG"
      switch_2 = JIG
      $ 1498 "Case 7"
      if (7 == switch_2):
        $ 1511 "Bottle"
        $ 1512 "'CHANGE THE REFERENCE TO THE FRAME TO MOVE IN'"
        # 'CHANGE THE REFERENCE TO THE FRAME TO MOVE IN'
        $ 1518 "If TASK.ID≟43"
        if (TASK.ID == 43):
          $ 1519 "Frame & Position Params"
          $ 1520 "FRM_Reference = CAM_LM_Bott"
          FRM_Reference = CAM_LM_Bott
          $ 1521 "PSE_T≔uLM_SS_PickPlc"
          global PSE_T=uLM_SS_PickPlc
          $ 1522 "PSE_A≔pose_trans(PSE_T, p[0,0,0.1,0,0,0])"
          global PSE_A= pose_trans (PSE_T, p[0,0,0.1,0,0,0])
          $ 1523 "PSE_R≔pose_add(PSE_T, p[0,0,0.1,0,0,0])"
          global PSE_R= pose_add (PSE_T, p[0,0,0.1,0,0,0])
        end
      end
    end
    $ 1530 "Additional check"
    $ 1531 "If  not is_reachable(FRM_Reference,[PSE_A,PSE_A_H,PSE_T,PSE_T_H,PSE_R,PSE_R_H])"
    if (  not  is_reachable(FRM_Reference,[PSE_A,PSE_A_H,PSE_T,PSE_T_H,PSE_R,PSE_R_H])):
      $ 1532 "Error"
      $ 1533 "set_error(ERROR_POSE_NOT_REACHABLE)"
      set_error(ERROR_POSE_NOT_REACHABLE)
      $ 1534 "Action≔0"
      global Action=0
    end
    $ 1535 "'=========='"
    # '=========='
    $ 1536 "Switch Action"
    switch_1 = Action
    $ 1537 "Case 1"
    if (1 == switch_1):
      $ 1538 "Pick"
      $ 1539 "Action_Info≔'pick object'"
      global Action_Info="pick object"
      $ 1540 "do_transition(pose_trans(FRM_Reference, PSE_T), keep_rxry=OBJ_Picked)"
      do_transition( pose_trans (FRM_Reference, PSE_T), keep_rxry=OBJ_Picked)
      $ 1541 "EOAT"
      $ 1542 "If  not OBJ_Picked"
      if (  not  OBJ_Picked):
        $ 1543 "rq_move_and_wait_mm(GRP_Open_Pos)"
         rq_move_and_wait_mm (GRP_Open_Pos)
      end
      $ 1544 "If PSE_A_H≠PSE_Z"
      if (PSE_A_H != PSE_Z):
        $ 1545 "If JNT_Q≠JNT_Z"
        if (JNT_Q != JNT_Z):
          $ 1546 "movej(get_inverse_kin(pose_trans(FRM_Reference, PSE_A_H), qnear=JNT_Q), r=0.050)"
          movej(get_inverse_kin( pose_trans (FRM_Reference, PSE_A_H), qnear=JNT_Q), r=0.050)
        else:
          $ 1547 "Else" "noBreak"
          $ 1548 "movej(pose_trans(FRM_Reference, PSE_A_H), r=0.050)"
          movej( pose_trans (FRM_Reference, PSE_A_H), r=0.050)
        end
      end
      $ 1549 "If PSE_A≠PSE_Z"
      if (PSE_A != PSE_Z):
        $ 1550 "If JNT_Q≠JNT_Z"
        if (JNT_Q != JNT_Z):
          $ 1551 "movej(get_inverse_kin(pose_trans(FRM_Reference, PSE_A), qnear=JNT_Q), r=0.020)"
          movej(get_inverse_kin( pose_trans (FRM_Reference, PSE_A), qnear=JNT_Q), r=0.020)
        else:
          $ 1552 "Else" "noBreak"
          $ 1553 "movej(pose_trans(FRM_Reference, PSE_A), r=0.020)"
          movej( pose_trans (FRM_Reference, PSE_A), r=0.020)
        end
      end
      $ 1554 "MoveL"
      $ 1555 "If PSE_T_H≠PSE_Z"
      if (PSE_T_H != PSE_Z):
        $ 1556 "PSE_T_H" "breakAfter"
        movel(pose_trans(FRM_Reference, PSE_T_H), a=0.5, v=0.4, r=0.01)
      end
      $ 1557 "PSE_T" "breakAfter"
      movel(pose_trans(FRM_Reference, PSE_T), a=0.08, v=0.12)
      $ 1558 "EOAT"
      $ 1559 "rq_set_force_norm(50)"
       rq_set_force_norm (50)
      $ 1560 "rq_close_and_wait()"
       rq_close_and_wait ()
      $ 1561 "OBJ_Picked≔rq_is_object_detected()"
      global OBJ_Picked= rq_is_object_detected ()
      $ 1562 "If  not OBJ_Picked"
      if (  not  OBJ_Picked):
        $ 1563 "set_error(ERROR_NO_OBJECT_TO_PICK)"
        set_error(ERROR_NO_OBJECT_TO_PICK)
      end
      $ 1564 "EXTT"
      $ 1565 "Switch JIG"
      switch_2 = JIG
      $ 1566 "Case 1"
      if (1 == switch_2):
        $ 1567 "3FG"
        $ 1568 "If OBJ_Picked"
        if (OBJ_Picked):
          $ 1569 "Set GRP_3F_Open=On"
          set_standard_digital_out(5, True)
        end
      end
      $ 1570 "If PSE_R_H≠PSE_Z"
      if (PSE_R_H != PSE_Z):
        $ 1571 "PSE_R" "breakAfter"
        movel(pose_trans(FRM_Reference, PSE_R), a=0.5, v=0.4, r=0.01)
        $ 1572 "PSE_R_H" "breakAfter"
        movel(pose_trans(FRM_Reference, PSE_R_H), a=0.5, v=0.4)
      else:
        $ 1573 "Else" "noBreak"
        $ 1574 "PSE_R" "breakAfter"
        movel(pose_trans(FRM_Reference, PSE_R), a=0.5, v=0.4)
      end
    elif (2 == switch_1):
      $ 1575 "Case 2"
    elif (3 == switch_1):
      $ 1617 "Case 3"
    elif (4 == switch_1):
      $ 1620 "Case 4"
    elif (5 == switch_1):
      $ 1623 "Case 5"
      $ 1624 "Pick the deepwell rack"
      # begin: URCap Program Node
      #   Source: SensoPart VISOR Robotic, 2.0.0, SensoPart Industriesensorik GmbH
      #   Type: VISOR Robotic App
      $ 1625 "VISOR Easy Pick"
      def visorFuncEasyPick_634681():
        # begin: URCap Program Node
        #   Source: SensoPart VISOR Robotic, 2.0.0, SensoPart Industriesensorik GmbH
        #   Type: Easy Pick Setup
        $ 1626 "# 1 Setup" "noBreak"
        local easyPickVisorId = 1
        local easyPickArmMounted = True
        local easyPickSetJob = True
        local easyPickJobName = "pick_rack"
        local easyPickAtImgAcq = False
        local easyPickImgAcqPose = FRM_Container_S
        # end: URCap Program Node
        # begin: URCap Program Node
        #   Source: SensoPart VISOR Robotic, 2.0.0, SensoPart Industriesensorik GmbH
        #   Type: Process
        $ 1627 "Process" "noBreak"
        local easyPickObjTaken = False
        local easyPickTrigger = False
        local easyPickPoseIdx = 0
        local easyPickPose = p[0,0,0,0,0,0]
        def easyPickFuncTrigger(visorId, setJob, jobName, arm):
        if (setJob):
          visor_changeJob(visorId, jobName, 6000)
        end
        if (arm):
          visor_trigger(visorId, 6000, "arm")
        else:
          visor_trigger(visorId, 6000)
        end
        global easyPickParts=visor_partsFound(visorId)
        visor_easyPickUpdate(visorId, "parts", visor_partsFound(visorId))
        return visor_getPose3d(visorId, 0)
      end
      while (not easyPickObjTaken):
        easyPickTrigger = (easyPickCount >= visor_partsFound(easyPickVisorId)) or (easyPickCount > 9) or (not visor_easyPickCheckIdent("efe41c", easyPickVisorId))
        if (easyPickTrigger):
          easyPickCount = 0
        end
        easyPickPoseIdx = easyPickCount
        easyPickPose = visor_getPose3d(easyPickVisorId, easyPickPoseIdx)
        visor_easyPickUpdate(easyPickVisorId, "counter", easyPickPoseIdx)
        # begin: URCap Program Node
        #   Source: SensoPart VISOR Robotic, 2.0.0, SensoPart Industriesensorik GmbH
        #   Type: Image Acquisition Pose
        $ 1628 "Image Acquisition Pose" "noBreak"
        if (easyPickTrigger):
          if (not easyPickAtImgAcq):
            movej(pose_trans(easyPickImgAcqPose,p[0.0000,0.0000,-0.0000,0.0000,0.0000,0.0000]),a=1.3963,v=1.0472,t=0.000000,r=0.000000)
            easyPickAtImgAcq = True
          end
          easyPickPose = easyPickFuncTrigger(easyPickVisorId, easyPickSetJob, easyPickJobName, easyPickArmMounted)
        end
        # end: URCap Program Node
        # begin: URCap Program Node
        #   Source: SensoPart VISOR Robotic, 2.0.0, SensoPart Industriesensorik GmbH
        #   Type: Object Detected
        $ 1629 "Object Detected" "noBreak"
        if (visor_partsFound(easyPickVisorId) > 0):
          $ 1630 "Open Gripper" "noBreak"
          # begin: URCap Program Node
          #   Source: Robotiq_Grippers, 1.8.4.4844, Robotiq Inc.
          #   Type: Gripper
          $ 1631 "Gripper Open (1)" "noBreak"
          if not(gripper_connected[0]):
            popup("Gripper 1 must be connected to run this program.", "No connection", False, True, True)
          end
          if not(rq_is_gripper_activated("1")):
            popup("Gripper 1 is not activated. Go to Installation tab > Gripper to activate it and run the program again.", "Not activated", False, True, True)
          end
          rq_set_pos_spd_for(0, 102, 77, "1")
          rq_wait_pos_spe_for_request(0, 102, 77, "1")
          rq_go_to("1")
          rq_wait("1")
          # end: URCap Program Node
          $ 1632 "MoveJ" "noBreak"
          $ 1633 "Waypoint_86" "noBreak"
          movej(get_inverse_kin(Waypoint_86_p, qnear=Waypoint_86_q), a=0.6981317007977318, v=0.5235987755982988)
          # begin: URCap Program Node
          #   Source: SensoPart VISOR Robotic, 2.0.0, SensoPart Industriesensorik GmbH
          #   Type: Approach Pose
          $ 1634 "Approach Pose" "noBreak"
          movej(pose_trans(easyPickPose,p[0.0000,0.0000,0.0500,0.0000,0.0000,0.0000]),a=0.6981,v=0.5236,t=0.000000,r=0.000000)
          # end: URCap Program Node
          # begin: URCap Program Node
          #   Source: SensoPart VISOR Robotic, 2.0.0, SensoPart Industriesensorik GmbH
          #   Type: Target Pose
          $ 1635 "Target Pose" "noBreak"
          movel(pose_trans(easyPickPose,p[0.0000,0.0000,-0.0000,0.0000,0.0000,0.0000]),a=0.2000,v=0.1200,t=0.000000,r=0.000000)
          # end: URCap Program Node
          $ 1636 "Close Gripper" "noBreak"
          # begin: URCap Program Node
          #   Source: Robotiq_Grippers, 1.8.4.4844, Robotiq Inc.
          #   Type: Gripper
          $ 1637 "Gripper Close (1)" "noBreak"
          if not(gripper_connected[0]):
            popup("Gripper 1 must be connected to run this program.", "No connection", False, True, True)
          end
          if not(rq_is_gripper_activated("1")):
            popup("Gripper 1 is not activated. Go to Installation tab > Gripper to activate it and run the program again.", "Not activated", False, True, True)
          end
          rq_set_pos_spd_for(255, 102, 77, "1")
          rq_wait_pos_spe_for_request(255, 102, 77, "1")
          rq_go_to("1")
          rq_wait("1")
          # end: URCap Program Node
          # begin: URCap Program Node
          #   Source: SensoPart VISOR Robotic, 2.0.0, SensoPart Industriesensorik GmbH
          #   Type: Exit Pose
          $ 1638 "Exit Pose" "noBreak"
          movel(pose_trans(easyPickPose,p[0.0000,0.0000,-0.0000,0.0000,0.0000,0.0000]),a=0.2000,v=0.1200,t=0.000000,r=0.000000)
          # end: URCap Program Node
          easyPickObjTaken = True
        end
        # end: URCap Program Node
        # begin: URCap Program Node
        #   Source: SensoPart VISOR Robotic, 2.0.0, SensoPart Industriesensorik GmbH
        #   Type: No Object Detected
        $ 1639 "No Object Detected" "noBreak"
        if (visor_partsFound(easyPickVisorId) < 1):
          $ 1640 "Popup: No Container detected" "noBreak"
          popup("No Container detected", "Message", False, False, blocking=True)
          else:
        end
        # end: URCap Program Node
      end
      easyPickCount = easyPickCount + 1
      visor_easyPickUpdate(easyPickVisorId, "counter", easyPickCount)
      visor_easyPickSetIdent("efe41c", easyPickVisorId)
      # end: URCap Program Node
    end
    visorFuncEasyPick_634681()
    # end: URCap Program Node
    $ 1641 "Wait: 2.0"
    sleep(2.0)
    $ 1642 "MoveJ"
    $ 1643 "Waypoint_16" "breakAfter"
    movej(get_inverse_kin(Waypoint_16_p, qnear=Waypoint_16_q), a=0.6981317007977318, v=0.3490658503988659)
    $ 1644 "Waypoint_87" "breakAfter"
    movej(get_inverse_kin(Waypoint_87_p, qnear=Waypoint_87_q), a=0.6981317007977318, v=0.3490658503988659)
    $ 1645 "Waypoint_89" "breakAfter"
    movej(get_inverse_kin(Waypoint_89_p, qnear=Waypoint_89_q), a=0.6981317007977318, v=0.3490658503988659)
    $ 1646 "MoveL"
    $ 1647 "Waypoint_90" "breakAfter"
    movel(Waypoint_90_p, a=0.6, v=0.12)
    # begin: URCap Program Node
    #   Source: Robotiq_Grippers, 1.8.4.4844, Robotiq Inc.
    #   Type: Gripper
    $ 1648 "Gripper Open (1)"
    if not(gripper_connected[0]):
      popup("Gripper 1 must be connected to run this program.", "No connection", False, True, True)
    end
    if not(rq_is_gripper_activated("1")):
      popup("Gripper 1 is not activated. Go to Installation tab > Gripper to activate it and run the program again.", "Not activated", False, True, True)
    end
    rq_set_pos_spd_for(0, 0, 0, "1")
    rq_wait_pos_spe_for_request(0, 0, 0, "1")
    rq_go_to("1")
    rq_wait("1")
    # end: URCap Program Node
    $ 1649 "Waypoint_89" "breakAfter"
    movel(Waypoint_89_p, a=0.6, v=0.12)
  elif (6 == switch_1):
    $ 1650 "Case 6"
    $ 1665 "offset≔p[0, 0.03, 0, 0, 0, 0]"
    global offset=p[0, 0.03, 0, 0, 0, 0]
    $ 1666 "Place the deepwell rack"
    # begin: URCap Program Node
    #   Source: SensoPart VISOR Robotic, 2.0.0, SensoPart Industriesensorik GmbH
    #   Type: VISOR Robotic App
    $ 1667 "VISOR Easy Pick"
    def visorFuncEasyPick_b634ba():
      # begin: URCap Program Node
      #   Source: SensoPart VISOR Robotic, 2.0.0, SensoPart Industriesensorik GmbH
      #   Type: Easy Pick Setup
      $ 1668 "# 1 Setup" "noBreak"
      local easyPickVisorId = 1
      local easyPickArmMounted = True
      local easyPickSetJob = True
      local easyPickJobName = "place_rack"
      local easyPickAtImgAcq = False
      local easyPickImgAcqPose = aq_rack1
      # end: URCap Program Node
      # begin: URCap Program Node
      #   Source: SensoPart VISOR Robotic, 2.0.0, SensoPart Industriesensorik GmbH
      #   Type: Process
      $ 1669 "Process" "noBreak"
      local easyPickObjTaken = False
      local easyPickTrigger = False
      local easyPickPoseIdx = 0
      local easyPickPose = p[0,0,0,0,0,0]
      def easyPickFuncTrigger(visorId, setJob, jobName, arm):
      if (setJob):
        visor_changeJob(visorId, jobName, 6000)
      end
      if (arm):
        visor_trigger(visorId, 6000, "arm")
      else:
        visor_trigger(visorId, 6000)
      end
      global easyPickParts=visor_partsFound(visorId)
      visor_easyPickUpdate(visorId, "parts", visor_partsFound(visorId))
      return visor_getPose3d(visorId, 0)
    end
    while (not easyPickObjTaken):
      easyPickTrigger = (easyPickCount >= visor_partsFound(easyPickVisorId)) or (easyPickCount > 9) or (not visor_easyPickCheckIdent("1b32aa", easyPickVisorId))
      if (easyPickTrigger):
        easyPickCount = 0
      end
      easyPickPoseIdx = easyPickCount
      easyPickPose = visor_getPose3d(easyPickVisorId, easyPickPoseIdx)
      visor_easyPickUpdate(easyPickVisorId, "counter", easyPickPoseIdx)
      # begin: URCap Program Node
      #   Source: SensoPart VISOR Robotic, 2.0.0, SensoPart Industriesensorik GmbH
      #   Type: Image Acquisition Pose
      $ 1670 "Image Acquisition Pose" "noBreak"
      if (easyPickTrigger):
        if (not easyPickAtImgAcq):
          movej(pose_trans(easyPickImgAcqPose,p[0.0000,0.0000,-0.0000,0.0000,0.0000,0.0000]),a=1.3963,v=1.0472,t=0.000000,r=0.000000)
          easyPickAtImgAcq = True
        end
        easyPickPose = easyPickFuncTrigger(easyPickVisorId, easyPickSetJob, easyPickJobName, easyPickArmMounted)
      end
      # end: URCap Program Node
      # begin: URCap Program Node
      #   Source: SensoPart VISOR Robotic, 2.0.0, SensoPart Industriesensorik GmbH
      #   Type: Object Detected
      $ 1671 "Object Detected" "noBreak"
      if (visor_partsFound(easyPickVisorId) > 0):
        $ 1672 "Open Gripper" "noBreak"
        # begin: URCap Program Node
        #   Source: Robotiq_Grippers, 1.8.4.4844, Robotiq Inc.
        #   Type: Gripper
        $ 1673 "Gripper Open (1)" "noBreak"
        if not(gripper_connected[0]):
          popup("Gripper 1 must be connected to run this program.", "No connection", False, True, True)
        end
        if not(rq_is_gripper_activated("1")):
          popup("Gripper 1 is not activated. Go to Installation tab > Gripper to activate it and run the program again.", "Not activated", False, True, True)
        end
        rq_set_pos_spd_for(0, 102, 77, "1")
        rq_wait_pos_spe_for_request(0, 102, 77, "1")
        rq_go_to("1")
        rq_wait("1")
        # end: URCap Program Node
        $ 1674 "MoveJ" "noBreak"
        $ 1675 "Waypoint_88" "noBreak"
        movej(get_inverse_kin(Waypoint_88_p, qnear=Waypoint_88_q), a=0.6981317007977318, v=0.5235987755982988)
        $ 1676 "Waypoint_87" "noBreak"
        movej(get_inverse_kin(Waypoint_87_p, qnear=Waypoint_87_q), a=0.6981317007977318, v=0.5235987755982988)
        $ 1677 "Waypoint_89" "noBreak"
        movej(get_inverse_kin(Waypoint_89_p, qnear=Waypoint_89_q), a=0.6981317007977318, v=0.5235987755982988)
        $ 1678 "MoveL" "noBreak"
        $ 1679 "Waypoint_90" "noBreak"
        movel(Waypoint_90_p, a=0.6, v=0.12)
        # begin: URCap Program Node
        #   Source: Robotiq_Grippers, 1.8.4.4844, Robotiq Inc.
        #   Type: Gripper
        $ 1680 "Gripper Close (1)" "noBreak"
        if not(gripper_connected[0]):
          popup("Gripper 1 must be connected to run this program.", "No connection", False, True, True)
        end
        if not(rq_is_gripper_activated("1")):
          popup("Gripper 1 is not activated. Go to Installation tab > Gripper to activate it and run the program again.", "Not activated", False, True, True)
        end
        rq_set_pos_spd_for(255, 0, 0, "1")
        rq_wait_pos_spe_for_request(255, 0, 0, "1")
        rq_go_to("1")
        rq_wait("1")
        # end: URCap Program Node
        $ 1681 "Waypoint_89" "noBreak"
        movel(Waypoint_89_p, a=0.6, v=0.12)
        $ 1685 "MoveJ" "noBreak"
        $ 1686 "Waypoint_94" "noBreak"
        movej(get_inverse_kin(Waypoint_94_p, qnear=Waypoint_94_q), a=1.3962634015954636, v=1.0471975511965976)
        $ 1687 "Waypoint_93" "noBreak"
        movej(get_inverse_kin(Waypoint_93_p, qnear=Waypoint_93_q), a=1.3962634015954636, v=1.0471975511965976)
        # begin: URCap Program Node
        #   Source: SensoPart VISOR Robotic, 2.0.0, SensoPart Industriesensorik GmbH
        #   Type: Approach Pose
        $ 1688 "Approach Pose" "noBreak"
        movej(pose_trans(easyPickPose,p[0.0000,0.0000,-0.0000,0.0000,0.0000,0.0000]),a=0.6981,v=0.5236,t=0.000000,r=0.000000)
        # end: URCap Program Node
        # begin: URCap Program Node
        #   Source: SensoPart VISOR Robotic, 2.0.0, SensoPart Industriesensorik GmbH
        #   Type: Target Pose
        $ 1689 "Target Pose" "noBreak"
        movel(pose_trans(easyPickPose,p[0.0000,0.0000,-0.0000,0.0000,0.0000,0.0000]),a=0.2000,v=0.1000,t=0.000000,r=0.000000)
        # end: URCap Program Node
        $ 1690 "Close Gripper" "noBreak"
        $ 1691 "current_pose≔get_actual_tcp_pose()" "noBreak"
        global current_pose= get_actual_tcp_pose ()
        $ 1692 "place_pose≔pose_trans(current_pose, offset)" "noBreak"
        global place_pose=pose_trans(current_pose, offset)
        $ 1693 "MoveJ" "noBreak"
        $ 1694 "place_pose" "noBreak"
        movej(place_pose, a=0.5235987755982988, v=0.3490658503988659)
        # begin: URCap Program Node
        #   Source: Robotiq_Grippers, 1.8.4.4844, Robotiq Inc.
        #   Type: Gripper
        $ 1695 "Gripper Open (1)" "noBreak"
        if not(gripper_connected[0]):
          popup("Gripper 1 must be connected to run this program.", "No connection", False, True, True)
        end
        if not(rq_is_gripper_activated("1")):
          popup("Gripper 1 is not activated. Go to Installation tab > Gripper to activate it and run the program again.", "Not activated", False, True, True)
        end
        rq_set_pos_spd_for(0, 0, 0, "1")
        rq_wait_pos_spe_for_request(0, 0, 0, "1")
        rq_go_to("1")
        rq_wait("1")
        # end: URCap Program Node
        # begin: URCap Program Node
        #   Source: SensoPart VISOR Robotic, 2.0.0, SensoPart Industriesensorik GmbH
        #   Type: Exit Pose
        $ 1696 "Exit Pose" "noBreak"
        movel(pose_trans(easyPickPose,p[0.0000,0.0000,-0.0000,0.0000,0.0000,0.0000]),a=0.2000,v=0.1200,t=0.000000,r=0.000000)
        # end: URCap Program Node
        easyPickObjTaken = True
      end
      # end: URCap Program Node
      # begin: URCap Program Node
      #   Source: SensoPart VISOR Robotic, 2.0.0, SensoPart Industriesensorik GmbH
      #   Type: No Object Detected
      $ 1697 "No Object Detected" "noBreak"
      if (visor_partsFound(easyPickVisorId) < 1):
        $ 1698 "Popup: No Container detected" "noBreak"
        popup("No Container detected", "Message", False, False, blocking=True)
        else:
      end
      # end: URCap Program Node
    end
    easyPickCount = easyPickCount + 1
    visor_easyPickUpdate(easyPickVisorId, "counter", easyPickCount)
    visor_easyPickSetIdent("1b32aa", easyPickVisorId)
    # end: URCap Program Node
